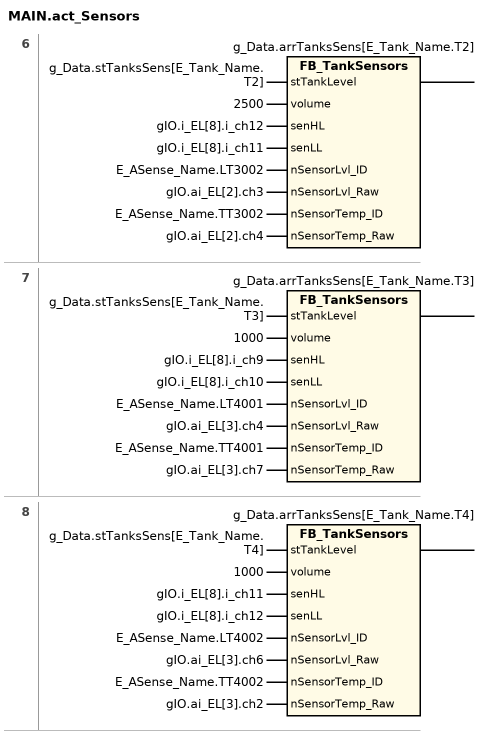
// NETWORK 6
g_Data.arrTanksSens[E_Tank_Name.T2](
    stTankLevel := g_Data.stTanksSens[E_Tank_Name.T2],
    volume := 2500,
    senHL := gIO.i_EL[8].i_ch12,
    senLL := gIO.i_EL[8].i_ch11,
    nSensorLvl_ID := E_ASense_Name.LT3002,
    nSensorLvl_Raw := gIO.ai_EL[2].ch3,
    nSensorTemp_ID := E_ASense_Name.TT3002,
    nSensorTemp_Raw := gIO.ai_EL[2].ch4); // FB_TankSensors

// NETWORK 7
g_Data.arrTanksSens[E_Tank_Name.T3](
    stTankLevel := g_Data.stTanksSens[E_Tank_Name.T3],
    volume := 1000,
    senHL := gIO.i_EL[8].i_ch9,
    senLL := gIO.i_EL[8].i_ch10,
    nSensorLvl_ID := E_ASense_Name.LT4001,
    nSensorLvl_Raw := gIO.ai_EL[3].ch4,
    nSensorTemp_ID := E_ASense_Name.TT4001,
    nSensorTemp_Raw := gIO.ai_EL[3].ch7); // FB_TankSensors

// NETWORK 8
g_Data.arrTanksSens[E_Tank_Name.T4](
    stTankLevel := g_Data.stTanksSens[E_Tank_Name.T4],
    volume := 1000,
    senHL := gIO.i_EL[8].i_ch11,
    senLL := gIO.i_EL[8].i_ch12,
    nSensorLvl_ID := E_ASense_Name.LT4002,
    nSensorLvl_Raw := gIO.ai_EL[3].ch6,
    nSensorTemp_ID := E_ASense_Name.TT4002,
    nSensorTemp_Raw := gIO.ai_EL[3].ch2); // FB_TankSensors
END_ACTION

ACTION act_SetAnalogSens_Test:
//set analog sensors setting only for the test. 
//Later this action should be deleted 
IF NOT bTesting THEN
	//Level
	g_AnalogSensor.stAnalogSensor[E_ASense_Name.LT1004].rawVal_Max:=14350;
	g_AnalogSensor.stAnalogSensor[E_ASense_Name.LT1004].rawVal_Min:=1270;
	g_AnalogSensor.stAnalogSensor[E_ASense_Name.LT1004].outVal_Max:=785;
	g_AnalogSensor.stAnalogSensor[E_ASense_Name.LT1004].outVal_Min:=0;
	g_AnalogSensor.stAnalogSensor[E_ASense_Name.LT1004].outOffset:=73;
	
	g_AnalogSensor.stAnalogSensor[E_ASense_Name.LT1003].rawVal_Max:=14350;
	g_AnalogSensor.stAnalogSensor[E_ASense_Name.LT1003].rawVal_Min:=1270;
	g_AnalogSensor.stAnalogSensor[E_ASense_Name.LT1003].outVal_Max:=785;
	g_AnalogSensor.stAnalogSensor[E_ASense_Name.LT1003].outVal_Min:=0;
	g_AnalogSensor.stAnalogSensor[E_ASense_Name.LT1003].outOffset:=73;
	
	g_AnalogSensor.stAnalogSensor[E_ASense_Name.LT1002].rawVal_Max:=14350;
	g_AnalogSensor.stAnalogSensor[E_ASense_Name.LT1002].rawVal_Min:=1270;
	g_AnalogSensor.stAnalogSensor[E_ASense_Name.LT1002].outVal_Max:=785;
	g_AnalogSensor.stAnalogSensor[E_ASense_Name.LT1002].outVal_Min:=0;
	g_AnalogSensor.stAnalogSensor[E_ASense_Name.LT1002].outOffset:=73;
	
	g_AnalogSensor.stAnalogSensor[E_ASense_Name.LT1001].rawVal_Max:=14350;
	g_AnalogSensor.stAnalogSensor[E_ASense_Name.LT1001].rawVal_Min:=1270;
	g_AnalogSensor.stAnalogSensor[E_ASense_Name.LT1001].outVal_Max:=785;
	g_AnalogSensor.stAnalogSensor[E_ASense_Name.LT1001].outVal_Min:=0;
	g_AnalogSensor.stAnalogSensor[E_ASense_Name.LT1001].outOffset:=73;
	
	//Flow
	g_AnalogSensor.stAnalogSensor[E_ASense_Name.FT1001].rawVal_Max:=10000;
	g_AnalogSensor.stAnalogSensor[E_ASense_Name.FT1001].rawVal_Min:=0;
	g_AnalogSensor.stAnalogSensor[E_ASense_Name.FT1001].outVal_Max:=306;
	g_AnalogSensor.stAnalogSensor[E_ASense_Name.FT1001].outVal_Min:=0;
	g_AnalogSensor.stAnalogSensor[E_ASense_Name.FT1001].outOffset:=0;
	
	g_AnalogSensor.stAnalogSensor[E_ASense_Name.FT1002].rawVal_Max:=10000;
	g_AnalogSensor.stAnalogSensor[E_ASense_Name.FT1002].rawVal_Min:=0;
	g_AnalogSensor.stAnalogSensor[E_ASense_Name.FT1002].outVal_Max:=306;
	g_AnalogSensor.stAnalogSensor[E_ASense_Name.FT1002].outVal_Min:=0;
	g_AnalogSensor.stAnalogSensor[E_ASense_Name.FT1002].outOffset:=0;
	
	////conductivity sensors
	g_AnalogSensor.stAnalogSensor[E_ASense_Name.CT1101].rawVal_Max:=14150;
	g_AnalogSensor.stAnalogSensor[E_ASense_Name.CT1101].rawVal_Min:=305;
	g_AnalogSensor.stAnalogSensor[E_ASense_Name.CT1101].outVal_Max:=14560;
	g_AnalogSensor.stAnalogSensor[E_ASense_Name.CT1101].outVal_Min:=346;
	g_AnalogSensor.stAnalogSensor[E_ASense_Name.CT1101].outOffset:=0;
	(*
	g_AnalogSensor.stAnalogSensor[E_ASense_Name.CT3101].rawVal_Max:=14150;
	g_AnalogSensor.stAnalogSensor[E_ASense_Name.CT3101].rawVal_Min:=305;
	g_AnalogSensor.stAnalogSensor[E_ASense_Name.CT3101].outVal_Max:=14560;
	g_AnalogSensor.stAnalogSensor[E_ASense_Name.CT3101].outVal_Min:=346;
	g_AnalogSensor.stAnalogSensor[E_ASense_Name.CT3101].outOffset:=0;
	*)
	//Temperature sensor
	g_AnalogSensor.stAnalogSensor[E_ASense_Name.TT1001].rawVal_Max:=7470;
	g_AnalogSensor.stAnalogSensor[E_ASense_Name.TT1001].rawVal_Min:=6400;
	g_AnalogSensor.stAnalogSensor[E_ASense_Name.TT1001].outVal_Max:=26;
	g_AnalogSensor.stAnalogSensor[E_ASense_Name.TT1001].outVal_Min:=20.9;
	g_AnalogSensor.stAnalogSensor[E_ASense_Name.TT1001].outOffset:=0;
	
	g_AnalogSensor.stAnalogSensor[E_ASense_Name.TT1002].rawVal_Max:=7470;
	g_AnalogSensor.stAnalogSensor[E_ASense_Name.TT1002].rawVal_Min:=6400;
	g_AnalogSensor.stAnalogSensor[E_ASense_Name.TT1002].outVal_Max:=26;
	g_AnalogSensor.stAnalogSensor[E_ASense_Name.TT1002].outVal_Min:=20.9;
	g_AnalogSensor.stAnalogSensor[E_ASense_Name.TT1002].outOffset:=0;
	
	g_AnalogSensor.stAnalogSensor[E_ASense_Name.TT1003].rawVal_Max:=7470;
	g_AnalogSensor.stAnalogSensor[E_ASense_Name.TT1003].rawVal_Min:=6400;
	g_AnalogSensor.stAnalogSensor[E_ASense_Name.TT1003].outVal_Max:=26;
	g_AnalogSensor.stAnalogSensor[E_ASense_Name.TT1003].outVal_Min:=20.9;
	g_AnalogSensor.stAnalogSensor[E_ASense_Name.TT1003].outOffset:=0;
	
	g_AnalogSensor.stAnalogSensor[E_ASense_Name.TT1004].rawVal_Max:=7470;
	g_AnalogSensor.stAnalogSensor[E_ASense_Name.TT1004].rawVal_Min:=6400;
	g_AnalogSensor.stAnalogSensor[E_ASense_Name.TT1004].outVal_Max:=26;
	g_AnalogSensor.stAnalogSensor[E_ASense_Name.TT1004].outVal_Min:=20.9;
	g_AnalogSensor.stAnalogSensor[E_ASense_Name.TT1004].outOffset:=0;
	
	g_AnalogSensor.stAnalogSensor[E_ASense_Name.TT1101].rawVal_Max:=7470;
	g_AnalogSensor.stAnalogSensor[E_ASense_Name.TT1101].rawVal_Min:=6400;
	g_AnalogSensor.stAnalogSensor[E_ASense_Name.TT1101].outVal_Max:=26;
	g_AnalogSensor.stAnalogSensor[E_ASense_Name.TT1101].outVal_Min:=20.9;
	g_AnalogSensor.stAnalogSensor[E_ASense_Name.TT1101].outOffset:=0;

	bTesting:=TRUE;
END_IF
END_ACTION

ACTION act_SetValves:
//Production tank
	//Tank1
	g_Data.arr_TankValves[1].valOutlet:=	E_Pis_Name.V3016;
	g_Data.arr_TankValves[1].valLine:=		E_Pis_Name.V3017;
	g_Data.arr_TankValves[1].valTriBlender:=E_Pis_Name.V3023;
	g_Data.arr_TankValves[1].valDrain:=		E_Pis_Name.V3024;
	g_Data.arr_TankValves[1].valCIP:=		E_Pis_Name.V3025;
	
	g_Data.arr_LineSourceValves[1].valTankA:=			E_Pis_Name.V3017;
	g_Data.arr_LineSourceValves[1].valTankB:=			E_Pis_Name.V3027;
	g_Data.arr_LineSourceValves[1].valTapWater:=		E_Pis_Name.V_Dummy_LSM_01;
	g_Data.arr_LineSourceValves[1].valTapWater_Drain:=	E_Pis_Name.V_Dummy_LSM_02;
	g_Data.arr_LineSourceValves[1].valTapWater_esle:=	E_Pis_Name.V_Dummy_LSM_05;
	g_Data.arr_LineSourceValves[1].valDrain:=			E_Pis_Name.V3018;
	g_Data.arr_LineSourceValves[1].valCIP:=				E_Pis_Name.V3019;
	g_Data.arr_LineSourceValves[1].valCIP_Sel:=			E_Pis_Name.V_Dummy_LSM_06;
	g_Data.arr_LineSourceValves[1].valBlockWater:=		E_Pis_Name.V_Dummy_LSM_03;
	g_Data.arr_LineSourceValves[1].valWaterSource:=		E_Pis_Name.V_Dummy_LSM_04;
	g_Data.arr_LineSourceValves[1].valWaterSource_Drain:=		E_Pis_Name.V_Dummy_LSM_07;
	
	g_Data.arr_TriBlenderSourceValves[1].valTankA:=				E_Pis_Name.V3023;
	g_Data.arr_TriBlenderSourceValves[1].valTankB:=				E_Pis_Name.V3028;
	g_Data.arr_TriBlenderSourceValves[1].valTapWater:=			E_Pis_Name.V_Dummy_TSM_01;
	g_Data.arr_TriBlenderSourceValves[1].valTapWater_Drain:=	E_Pis_Name.V_Dummy_TSM_02;
	g_Data.arr_TriBlenderSourceValves[1].valTapWater_esle:=		E_Pis_Name.V_Dummy_TSM_03;
	g_Data.arr_TriBlenderSourceValves[1].valDrain:=				E_Pis_Name.V3021;
	g_Data.arr_TriBlenderSourceValves[1].valCIP:=				E_Pis_Name.V3022;
	g_Data.arr_TriBlenderSourceValves[1].valCIP_Sel:=			E_Pis_Name.V3020;
	g_Data.arr_TriBlenderSourceValves[1].valBlockWater:=		E_Pis_Name.V3014;
	g_Data.arr_TriBlenderSourceValves[1].valWaterSource:=		E_Pis_Name.V3113;
	g_Data.arr_TriBlenderSourceValves[1].valWaterSource_Drain:=	E_Pis_Name.V2211;
	
	g_Data.arr_LineTargetValves[1].valTankA:=			E_Pis_Name.V_Dummy_01;//0;
	g_Data.arr_LineTargetValves[1].valTankB:=			E_Pis_Name.V_Dummy_02;//0;
	g_Data.arr_LineTargetValves[1].valDrain:=			E_Pis_Name.V_Dummy_03;//0;
	g_Data.arr_LineTargetValves[1].valCIP:=				E_Pis_Name.V_Dummy_04;//0;
	g_Data.arr_LineTargetValves[1].valTankA_Pipe:=		E_Pis_Name.V_Dummy_05;//0;
	g_Data.arr_LineTargetValves[1].valTankB_Pipe:=		E_Pis_Name.V_Dummy_06;//0;
	
	g_Data.arr_fbTriBlenderTargetValves[1].valTankA:=	E_Pis_Name.V3004;
	g_Data.arr_fbTriBlenderTargetValves[1].valTankB:=	E_Pis_Name.V3010;
	g_Data.arr_fbTriBlenderTargetValves[1].valDrain:=	E_Pis_Name.V3008;
	g_Data.arr_fbTriBlenderTargetValves[1].valCIP:=		E_Pis_Name.V3009;
	g_Data.arr_fbTriBlenderTargetValves[1].valTankA_Pipe:=		E_Pis_Name.v3041;
	g_Data.arr_fbTriBlenderTargetValves[1].valTankB_Pipe:=		E_Pis_Name.v3040;
	
	//Tank2
	g_Data.arr_TankValves[2].valOutlet:=	E_Pis_Name.V3015;
	g_Data.arr_TankValves[2].valLine:=		E_Pis_Name.V3027;
	g_Data.arr_TankValves[2].valTriBlender:=E_Pis_Name.V3028;
	g_Data.arr_TankValves[2].valDrain:=		E_Pis_Name.V3029;
	g_Data.arr_TankValves[2].valCIP:=		E_Pis_Name.V3030;
	
	g_Data.arr_LineSourceValves[2].valTankA:=			E_Pis_Name.V3017;
	g_Data.arr_LineSourceValves[2].valTankB:=			E_Pis_Name.V3027;
	g_Data.arr_LineSourceValves[2].valTapWater:=		E_Pis_Name.V_Dummy_LSM_01;
	g_Data.arr_LineSourceValves[2].valTapWater_Drain:=	E_Pis_Name.V_Dummy_LSM_02;
	g_Data.arr_LineSourceValves[2].valTapWater_esle:=	E_Pis_Name.V_Dummy_LSM_05;
	g_Data.arr_LineSourceValves[2].valDrain:=			E_Pis_Name.V3018;
	g_Data.arr_LineSourceValves[2].valCIP:=				E_Pis_Name.V3019;
	g_Data.arr_LineSourceValves[2].valCIP_Sel:=			E_Pis_Name.V_Dummy_LSM_06;
	g_Data.arr_LineSourceValves[2].valBlockWater:=		E_Pis_Name.V_Dummy_LSM_03;
	g_Data.arr_LineSourceValves[2].valWaterSource:=		E_Pis_Name.V_Dummy_LSM_04;
	g_Data.arr_LineSourceValves[2].valWaterSource_Drain:=		E_Pis_Name.V_Dummy_LSM_07;
	
	
	g_Data.arr_TriBlenderSourceValves[2].valTankA:=				E_Pis_Name.V3023;
	g_Data.arr_TriBlenderSourceValves[2].valTankB:=				E_Pis_Name.V3028;
	g_Data.arr_TriBlenderSourceValves[2].valTapWater:=			E_Pis_Name.V_Dummy_TSM_01;
	g_Data.arr_TriBlenderSourceValves[2].valTapWater_Drain:=	E_Pis_Name.V_Dummy_TSM_02;
	g_Data.arr_TriBlenderSourceValves[2].valTapWater_esle:=		E_Pis_Name.V_Dummy_TSM_03;
	g_Data.arr_TriBlenderSourceValves[2].valDrain:=				E_Pis_Name.V3021;
	g_Data.arr_TriBlenderSourceValves[2].valCIP:=				E_Pis_Name.V3022;
	g_Data.arr_TriBlenderSourceValves[2].valCIP_Sel:=			E_Pis_Name.V3020;
	g_Data.arr_TriBlenderSourceValves[2].valBlockWater:=		E_Pis_Name.V3014;
	g_Data.arr_TriBlenderSourceValves[2].valWaterSource:=		E_Pis_Name.V3113;
	g_Data.arr_TriBlenderSourceValves[2].valWaterSource_Drain:=	E_Pis_Name.V2211;
	
	g_Data.arr_LineTargetValves[2].valTankA:=			E_Pis_Name.V_Dummy_01;//0;
	g_Data.arr_LineTargetValves[2].valTankB:=			E_Pis_Name.V_Dummy_02;//0;
	g_Data.arr_LineTargetValves[2].valDrain:=			E_Pis_Name.V_Dummy_03;//0;
	g_Data.arr_LineTargetValves[2].valCIP:=				E_Pis_Name.V_Dummy_04;//0;
	g_Data.arr_LineTargetValves[2].valTankA_Pipe:=		E_Pis_Name.V_Dummy_05;//0;
	g_Data.arr_LineTargetValves[2].valTankB_Pipe:=		E_Pis_Name.V_Dummy_06;//0;	
	
	(*
	g_Data.arr_LineTargetValves[2].valTankA:=			E_Pis_Name.V_Dummy_07;//0;
	g_Data.arr_LineTargetValves[2].valTankB:=			E_Pis_Name.V_Dummy_08;//0;
	g_Data.arr_LineTargetValves[2].valDrain:=			E_Pis_Name.V_Dummy_09;//0;
	g_Data.arr_LineTargetValves[2].valCIP:=				E_Pis_Name.V_Dummy_10;//0;
	g_Data.arr_LineTargetValves[2].valTankA_Pipe:=		E_Pis_Name.V_Dummy_11;//0;
	g_Data.arr_LineTargetValves[2].valTankB_Pipe:=		E_Pis_Name.V_Dummy_12;//0;
	*)
	
	g_Data.arr_fbTriBlenderTargetValves[2].valTankA:=			E_Pis_Name.V3004;
	g_Data.arr_fbTriBlenderTargetValves[2].valTankB:=			E_Pis_Name.V3010;
	g_Data.arr_fbTriBlenderTargetValves[2].valDrain:=			E_Pis_Name.V3008;
	g_Data.arr_fbTriBlenderTargetValves[2].valCIP:=				E_Pis_Name.V3009;
	g_Data.arr_fbTriBlenderTargetValves[2].valTankA_Pipe:=		E_Pis_Name.V3041;
	g_Data.arr_fbTriBlenderTargetValves[2].valTankB_Pipe:=		E_Pis_Name.V3040;
	
	//Tank3
	g_Data.arr_TankValves[3].valOutlet:=	E_Pis_Name.V4016;
	g_Data.arr_TankValves[3].valLine:=		E_Pis_Name.V4017;
	g_Data.arr_TankValves[3].valTriBlender:=E_Pis_Name.V4023;
	g_Data.arr_TankValves[3].valDrain:=		E_Pis_Name.V4024;
	g_Data.arr_TankValves[3].valCIP:=		E_Pis_Name.V4025;
	
	g_Data.arr_LineSourceValves[3].valTankA:=			E_Pis_Name.V4017;
	g_Data.arr_LineSourceValves[3].valTankB:=			E_Pis_Name.V4027;
	g_Data.arr_LineSourceValves[3].valTapWater:=		E_Pis_Name.V2115;
	g_Data.arr_LineSourceValves[3].valTapWater_Drain:=	E_Pis_Name.V2117;
	g_Data.arr_LineSourceValves[3].valTapWater_esle:=	E_Pis_Name.V2116;
	g_Data.arr_LineSourceValves[3].valDrain:=			E_Pis_Name.V4018;
	g_Data.arr_LineSourceValves[3].valCIP:=				E_Pis_Name.V4019;
	g_Data.arr_LineSourceValves[3].valCIP_Sel:=			E_Pis_Name.V_Dummy_LSC_01;
	g_Data.arr_LineSourceValves[3].valBlockWater:=		E_Pis_Name.V_Dummy_LSC_02;
	g_Data.arr_LineSourceValves[3].valWaterSource:=		E_Pis_Name.V_Dummy_LSC_03;
	g_Data.arr_LineSourceValves[3].valWaterSource_Drain:=		E_Pis_Name.V_Dummy_LSC_04;
	
	g_Data.arr_TriBlenderSourceValves[3].valTankA:=				E_Pis_Name.V4023;
	g_Data.arr_TriBlenderSourceValves[3].valTankB:=				E_Pis_Name.V4028;
	g_Data.arr_TriBlenderSourceValves[3].valTapWater:=			E_Pis_Name.V2116;
	g_Data.arr_TriBlenderSourceValves[3].valTapWater_Drain:=	E_Pis_Name.V2117;
	g_Data.arr_TriBlenderSourceValves[3].valTapWater_esle:=		E_Pis_Name.V2115;
	g_Data.arr_TriBlenderSourceValves[3].valDrain:=				E_Pis_Name.V4021;
	g_Data.arr_TriBlenderSourceValves[3].valCIP:=				E_Pis_Name.V4022;
	g_Data.arr_TriBlenderSourceValves[3].valCIP_Sel:=			E_Pis_Name.V4020;
	g_Data.arr_TriBlenderSourceValves[3].valBlockWater:=		E_Pis_Name.V4014;
	g_Data.arr_TriBlenderSourceValves[3].valWaterSource:=		E_Pis_Name.V2114;
	g_Data.arr_TriBlenderSourceValves[3].valWaterSource_Drain:=	E_Pis_Name.V2112;
	
	g_Data.arr_LineTargetValves[3].valTankA:=	E_Pis_Name.V4034;
	g_Data.arr_LineTargetValves[3].valTankB:=	E_Pis_Name.V4033;
	g_Data.arr_LineTargetValves[3].valDrain:=	E_Pis_Name.V4035;
	g_Data.arr_LineTargetValves[3].valCIP:=		E_Pis_Name.V4036;
	g_Data.arr_LineTargetValves[3].valTankA_Pipe:=		E_Pis_Name.V4041;
	g_Data.arr_LineTargetValves[3].valTankB_Pipe:=		E_Pis_Name.V4040;
	
	g_Data.arr_fbTriBlenderTargetValves[3].valTankA:=	E_Pis_Name.V4004;
	g_Data.arr_fbTriBlenderTargetValves[3].valTankB:=	E_Pis_Name.V4010;
	g_Data.arr_fbTriBlenderTargetValves[3].valDrain:=	E_Pis_Name.V4008;
	g_Data.arr_fbTriBlenderTargetValves[3].valCIP:=		E_Pis_Name.V4009;
	g_Data.arr_fbTriBlenderTargetValves[3].valTankA_Pipe:=		E_Pis_Name.V4041;
	g_Data.arr_fbTriBlenderTargetValves[3].valTankB_Pipe:=		E_Pis_Name.V4040;
	
	//Tank4
	g_Data.arr_TankValves[4].valOutlet:=	E_Pis_Name.V4015;
	g_Data.arr_TankValves[4].valLine:=		E_Pis_Name.V4027;
	g_Data.arr_TankValves[4].valTriBlender:=E_Pis_Name.V4028;
	g_Data.arr_TankValves[4].valDrain:=		E_Pis_Name.V4029;
	g_Data.arr_TankValves[4].valCIP:=		E_Pis_Name.V4030;
	
	g_Data.arr_LineSourceValves[4].valTankA:=			E_Pis_Name.V4017;
	g_Data.arr_LineSourceValves[4].valTankB:=			E_Pis_Name.V4027;
	g_Data.arr_LineSourceValves[4].valTapWater:=		E_Pis_Name.V2115;
	g_Data.arr_LineSourceValves[4].valTapWater_Drain:=	E_Pis_Name.V2117;
	g_Data.arr_LineSourceValves[4].valTapWater_esle:=	E_Pis_Name.V2116;
	g_Data.arr_LineSourceValves[4].valDrain:=			E_Pis_Name.V4018;
	g_Data.arr_LineSourceValves[4].valCIP:=				E_Pis_Name.V4019;
	g_Data.arr_LineSourceValves[4].valCIP_Sel:=			E_Pis_Name.V_Dummy_LSC_01;
	g_Data.arr_LineSourceValves[4].valBlockWater:=		E_Pis_Name.V_Dummy_LSC_02;
	g_Data.arr_LineSourceValves[4].valWaterSource:=		E_Pis_Name.V_Dummy_LSC_03;
	g_Data.arr_LineSourceValves[4].valWaterSource_Drain:=		E_Pis_Name.V_Dummy_LSC_04;
	
	g_Data.arr_TriBlenderSourceValves[4].valTankA:=				E_Pis_Name.V4023;
	g_Data.arr_TriBlenderSourceValves[4].valTankB:=				E_Pis_Name.V4028;
	g_Data.arr_TriBlenderSourceValves[4].valTapWater:=			E_Pis_Name.V2116;
	g_Data.arr_TriBlenderSourceValves[4].valTapWater_Drain:=	E_Pis_Name.V2117;
	g_Data.arr_TriBlenderSourceValves[4].valTapWater_esle:=		E_Pis_Name.V2115;
	g_Data.arr_TriBlenderSourceValves[4].valDrain:=				E_Pis_Name.V4021;
	g_Data.arr_TriBlenderSourceValves[4].valCIP:=				E_Pis_Name.V4022;
	g_Data.arr_TriBlenderSourceValves[4].valCIP_Sel:=			E_Pis_Name.V4020;
	g_Data.arr_TriBlenderSourceValves[4].valBlockWater:=		E_Pis_Name.V4014;
	g_Data.arr_TriBlenderSourceValves[4].valWaterSource:=		E_Pis_Name.V2114;
	g_Data.arr_TriBlenderSourceValves[4].valWaterSource_Drain:=	E_Pis_Name.V2112;
	
	g_Data.arr_LineTargetValves[4].valTankA:=	E_Pis_Name.V4034;
	g_Data.arr_LineTargetValves[4].valTankB:=	E_Pis_Name.V4033;
	g_Data.arr_LineTargetValves[4].valDrain:=	E_Pis_Name.V4035;
	g_Data.arr_LineTargetValves[4].valCIP:=		E_Pis_Name.V4036;
	g_Data.arr_LineTargetValves[4].valTankA_Pipe:=		E_Pis_Name.V4041;
	g_Data.arr_LineTargetValves[4].valTankB_Pipe:=		E_Pis_Name.V4040;
	
	g_Data.arr_fbTriBlenderTargetValves[4].valTankA:=	E_Pis_Name.V4004;
	g_Data.arr_fbTriBlenderTargetValves[4].valTankB:=	E_Pis_Name.V4010;
	g_Data.arr_fbTriBlenderTargetValves[4].valDrain:=	E_Pis_Name.V4008;
	g_Data.arr_fbTriBlenderTargetValves[4].valCIP:=		E_Pis_Name.V4009;
	g_Data.arr_fbTriBlenderTargetValves[4].valTankA_Pipe:=		E_Pis_Name.V4041;
	g_Data.arr_fbTriBlenderTargetValves[4].valTankB_Pipe:=		E_Pis_Name.V4040;
END_ACTION

METHOD m_TankConus_Level_Calculation : REAL
VAR_INPUT
	raw: REAL;

END_VAR
VAR
	kConus: REAL:=0.00000002149 ;
END_VAR
IF raw<1230 THEN;
	//m_TankConus_Level_Calculation:=kConus*raw^3;
ELSE;
	m_TankConus_Level_Calculation:=raw;
END_IF
END_METHOD

METHOD mElementList_SetName : BOOL
VAR_INPUT
END_VAR

VAR
	eASense_Name: E_ASense_Name;
	eProcCntrl: E_ProcessControl_Name;
END_VAR
FOR eASense_Name:=0 TO E_ASense_Name.last DO
	arAnalogSensorNameList[eASense_Name]:=TO_STRING(eASense_Name);
END_FOR

FOR eProcCntrl:=0 TO E_ProcessControl_Name.eProcCntrl_Last DO
	arr_ProcCntrl_NameList[eProcCntrl]:=TO_STRING(eProcCntrl);
	g_ProcControl.arr_stProcCntrl[eProcCntrl].idName:=TO_STRING(eProcCntrl);
END_FOR
END_METHOD

END_PROGRAM

// ---- 03 Project/40 Misc/FB_OpenClose_Vlave.TcPOU
FUNCTION_BLOCK FB_OpenClose_Vlave
VAR_INPUT
	val_AfterPump	: E_Pis_Name;
	Pump_ID			: E_Pump_List:=E_Pump_List.eNotSelected;
END_VAR
VAR_OUTPUT
END_VAR
VAR
	stPist	: REFERENCE TO ST_Piston;
	stPump	: REFERENCE TO ST_Pump	;
	bOneTime	:	BOOL	;
END_VAR

act_SetReference();

IF (stPump.bRun_Auto OR stPump.bRun_Man) THEN
	bOneTime:=FALSE;
	IF NOT stPist.st_Open THEN
		stPist.req_Open:=TRUE;
	END_IF
ELSE
	IF NOT stPist.st_Close AND NOT bOneTime THEN
		stPist.req_Close:=TRUE;
		bOneTime:=TRUE;
	END_IF
END_IF

ACTION act_SetReference:
stPist REF= stPis[val_AfterPump];
stPump REF= g_Pump.arr_st_Pump[Pump_ID];
END_ACTION

END_FUNCTION_BLOCK

// ---- 00 Library/00-General/TimeAndDate/prg_RealClock.TcPOU
PROGRAM prg_RealClock
VAR

(* Real Time Clock *)
(*	dtRealTime				: DATE_AND_TIME;
	sRealTime				: STRING[22];	
	stSystemTime			: TimeStruct;
	stSystemTime_Empty		: TimeStruct;
	sTime					: STRING[20];
	sDate					: STRING[20];
	sTimeWithMicroSec		: STRING[40];*)

	syncTimer 	: TON;
	fbGetLocalTime 	: NT_GetTime;
	fbRTC_EX2 	: RTC_EX2;
	presetTime 	: TimeStruct;
	syncTrigger 	: F_TRIG;
	bBusy 		: BOOL;
	bError 		: BOOL;
	nErrID 		: UDINT;
	temp1: DATE;
	temp2: TOD;
	NetId :STRING :='';
	bValid_RTCEX2 	: BOOL;
	nMicroseconds 	: DWORD;
	r_trigTrigger: R_TRIG;
	sRealTime_Date	 :STRING(25);
	
	bStartTime: BOOL;
	stStart: TimeStruct;
	sDelta: STRING;
	ton_OneMinuteCount: TON;
END_VAR

(*--------->Set Plc Clock<----------------*)

dtRealTime:=SYSTEMTIME_TO_DT(stSystemTime);
sRealTime:= DT_TO_STRING(dtRealTime);
sRealTime_Date:= DT_TO_STRING(dtRealTime);
sRealTime_Date:=right(sRealTime_Date,19);
temp1:=DT_TO_DATE(dtRealTime);
temp2:=DT_TO_TOD(dtRealTime);
sDate:=DATE_TO_STRING(temp1);
sDate:=DELETE(sDate,2,1);


sTime:=TOD_TO_STRING(temp2);
sTime:=DELETE(sTime,4,1);

sDateTime:=CONCAT(sDate,' ');
sDateTime:=CONCAT(sDateTime,sTime);

sTimeWithMicroSec:=CONCAT(sTime,'.');
sTimeWithMicroSec:=CONCAT(sTimeWithMicroSec,DWORD_TO_STRING(nMicroseconds));




	syncTimer(IN:=NOT SyncTimer.Q , PT:=T#100ms , Q=> , ET=> );
(*r_trigTrigger(CLK:=q_Trigger);*)
	fbGetLocalTime(
		NETID:='' ,
		START:=syncTimer.Q,
		(*START:=r_trigTrigger.Q,*)
		TMOUT:=T#5s ,
		BUSY=>bBusy ,
		ERR=>bError ,
		ERRID=>nErrId ,
		TIMESTR=>presetTime );

	(*syncTrigger(CLK:=NOT bBusy*)
	syncTrigger(CLK:= bBusy
					 AND NOT bError , Q=> );
	fbRTC_EX2(
		EN:=syncTrigger.Q ,
		PDT:=presetTime ,
		PMICRO:=0 ,
		Q=>bValid_RTCEX2 ,
		CDT=>stSystemTime ,
		CMICRO=>nMicroseconds );
		
act_TestDelta();	

ton_OneMinuteCount(PT:=T#1m, IN:=NOT ton_OneMinuteCount.Q);

ACTION act_TestDelta:
IF bStartTime THEN;
	bStartTime:=FALSE;
	stStart:=stSystemTime;
END_IF

sDelta:= m_DeltaTime(stStartTime:=stStart);
END_ACTION

METHOD m_DeltaTime : STRING
VAR_INPUT
	stStartTime  : TimeStruct;
END_VAR
VAR
	tDelta: TIME;
	dtDelta: DATE_AND_TIME;
	todDelta: TOD;


END_VAR
tDelta:=TO_TIME(SYSTEMTIME_TO_DT(stSystemTime)-SYSTEMTIME_TO_DT(stStartTime));

m_DeltaTime:=mTime_to_String_HMI(tInputTime:=tDelta,iSecondDisplay:=FALSE);

(*old
todDelta:=TIME_TO_TOD(tDelta);
m_DeltaTime:=TOD_TO_STRING(todDelta);
m_DeltaTime:=DELETE(m_DeltaTime,4,1);
//dtDelta:=TO_DT(SYSTEMTIME_TO_DT(stSystemTime)-SYSTEMTIME_TO_DT(stStartTime));
//m_DeltaTime:=TIME_TO_STRING(dtDelta);
*)
END_METHOD

METHOD mTime_to_String_HMI : STRING
VAR_INPUT
    tInputTime 		: TIME; // TIME type, stored internally as LTIME (ms)
	iSecondDisplay	: BOOL;
END_VAR
VAR
    nTotalSeconds : UDINT;
    nTotalHours : UDINT;
    nMinutes : UDINT;
    nSeconds : UDINT;
    sFormatted : STRING(20);
END_VAR
// Convert TIME to total seconds
nTotalSeconds := TO_UDINT(tInputTime) / 1000;

// Extract minutes and seconds
nMinutes := nTotalSeconds / 60;
nSeconds := nTotalSeconds MOD 60;

// Convert to total hours
nTotalHours := nMinutes / 60;
nMinutes := nMinutes MOD 60;

// Format output as HHHH:MM:SS (e.g., 0123:45:56)
sFormatted := CONCAT(UDINT_TO_STRING(nTotalHours),'h:');
IF nMinutes < 10 THEN
    sFormatted := CONCAT(sFormatted, '0');
END_IF
sFormatted := CONCAT(sFormatted, UDINT_TO_STRING(nMinutes));
sFormatted := CONCAT(sFormatted, 'm');

IF iSecondDisplay THEN;
	sFormatted := CONCAT(sFormatted, ':');
	IF nSeconds < 10 THEN
		sFormatted := CONCAT(sFormatted, '0');
	END_IF
	sFormatted := CONCAT(sFormatted, UDINT_TO_STRING(nSeconds));
	sFormatted := CONCAT(sFormatted, 's');	
END_IF

// Return formatted string
mTime_to_String_HMI := sFormatted;
END_METHOD

END_PROGRAM

// ---- 01 Instance/01 Piston/prg_Piston.TcPOU
PROGRAM prg_Piston
VAR
	fbPiston: FB_Piston;
	stPiston: ST_Piston;

	bPis_Next_P: BOOL;
	bPis_Next_N: BOOL;

	

	
	TON_0: TON;
	TON_1: TON;
	TON_2: TON;
	TON_3: TON;
	TON_4: TON;
	TON_5: TON;	
	i: INT;
END_VAR

act_InterLock();
act_Call_list_TanksMarinade();
act_Call_list_TanksColor();
act_Call_list_TanksCoolant();
act_Call_List_LineSource();
act_Call_List_LineTarget();
act_Call_list_CIP_SourceNTarget();
act_Call_list_CIP_Client();
act_Call_list_CIP_Tanks();
act_Call_list_Water();
act_Call_list_TriBlender_Selector();


IF bPis_Next_P THEN;
	m_Get_Next_P(iSel:=iPis_sel);
	bPis_Next_P:=FALSE;
END_IF

IF bPis_Next_N THEN;
	m_Get_Next_N(iSel:=iPis_sel);
	bPis_Next_N:=FALSE;
END_IF

FOR i:=0 TO E_Pis_Name.last DO
	ePisNameList:=i;
	arPisNameList[i]:=TO_STRING(ePisNameList);
END_FOR

ACTION act_Call_list_CIP_Client:
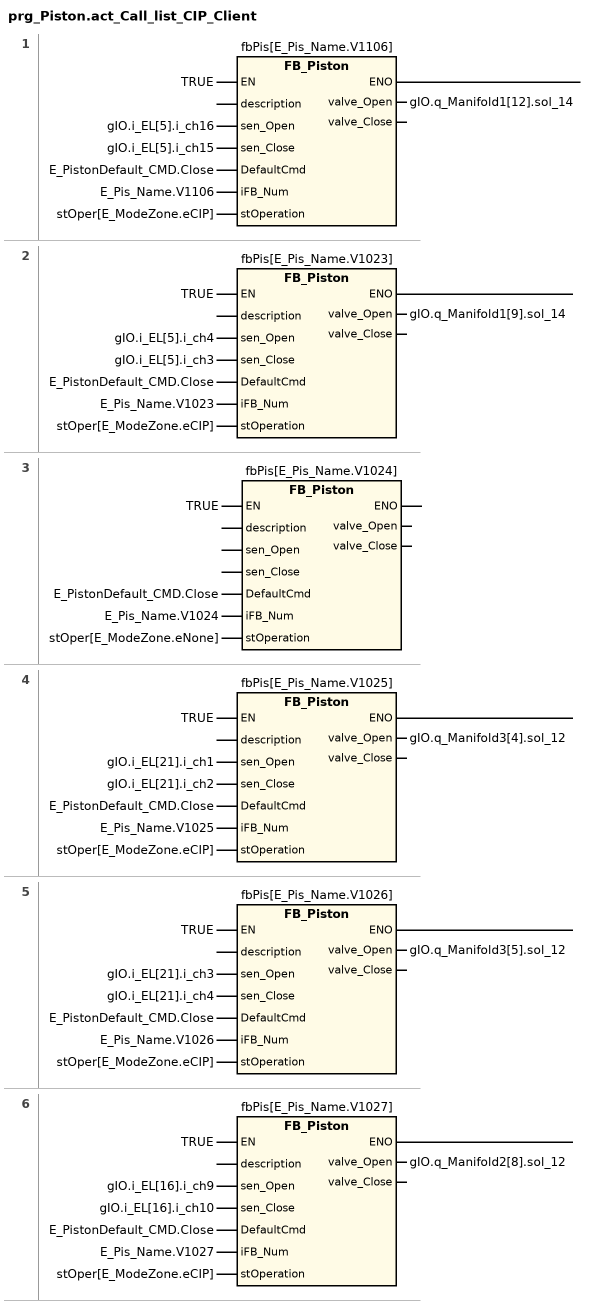
// NETWORK 1
fbPis[E_Pis_Name.V1106](
    sen_Open := gIO.i_EL[5].i_ch16,
    sen_Close := gIO.i_EL[5].i_ch15,
    DefaultCmd := E_PistonDefault_CMD.Close,
    iFB_Num := E_Pis_Name.V1106,
    stOperation := stOper[E_ModeZone.eCIP],
    valve_Open => gIO.q_Manifold1[12].sol_14); // FB_Piston

// NETWORK 2
fbPis[E_Pis_Name.V1023](
    sen_Open := gIO.i_EL[5].i_ch4,
    sen_Close := gIO.i_EL[5].i_ch3,
    DefaultCmd := E_PistonDefault_CMD.Close,
    iFB_Num := E_Pis_Name.V1023,
    stOperation := stOper[E_ModeZone.eCIP],
    valve_Open => gIO.q_Manifold1[9].sol_14); // FB_Piston

// NETWORK 3
fbPis[E_Pis_Name.V1024](
    DefaultCmd := E_PistonDefault_CMD.Close,
    iFB_Num := E_Pis_Name.V1024,
    stOperation := stOper[E_ModeZone.eNone]); // FB_Piston

// NETWORK 4
fbPis[E_Pis_Name.V1025](
    sen_Open := gIO.i_EL[21].i_ch1,
    sen_Close := gIO.i_EL[21].i_ch2,
    DefaultCmd := E_PistonDefault_CMD.Close,
    iFB_Num := E_Pis_Name.V1025,
    stOperation := stOper[E_ModeZone.eCIP],
    valve_Open => gIO.q_Manifold3[4].sol_12); // FB_Piston

// NETWORK 5
fbPis[E_Pis_Name.V1026](
    sen_Open := gIO.i_EL[21].i_ch3,
    sen_Close := gIO.i_EL[21].i_ch4,
    DefaultCmd := E_PistonDefault_CMD.Close,
    iFB_Num := E_Pis_Name.V1026,
    stOperation := stOper[E_ModeZone.eCIP],
    valve_Open => gIO.q_Manifold3[5].sol_12); // FB_Piston

// NETWORK 6
fbPis[E_Pis_Name.V1027](
    sen_Open := gIO.i_EL[16].i_ch9,
    sen_Close := gIO.i_EL[16].i_ch10,
    DefaultCmd := E_PistonDefault_CMD.Close,
    iFB_Num := E_Pis_Name.V1027,
    stOperation := stOper[E_ModeZone.eCIP],
    valve_Open => gIO.q_Manifold2[8].sol_12); // FB_Piston

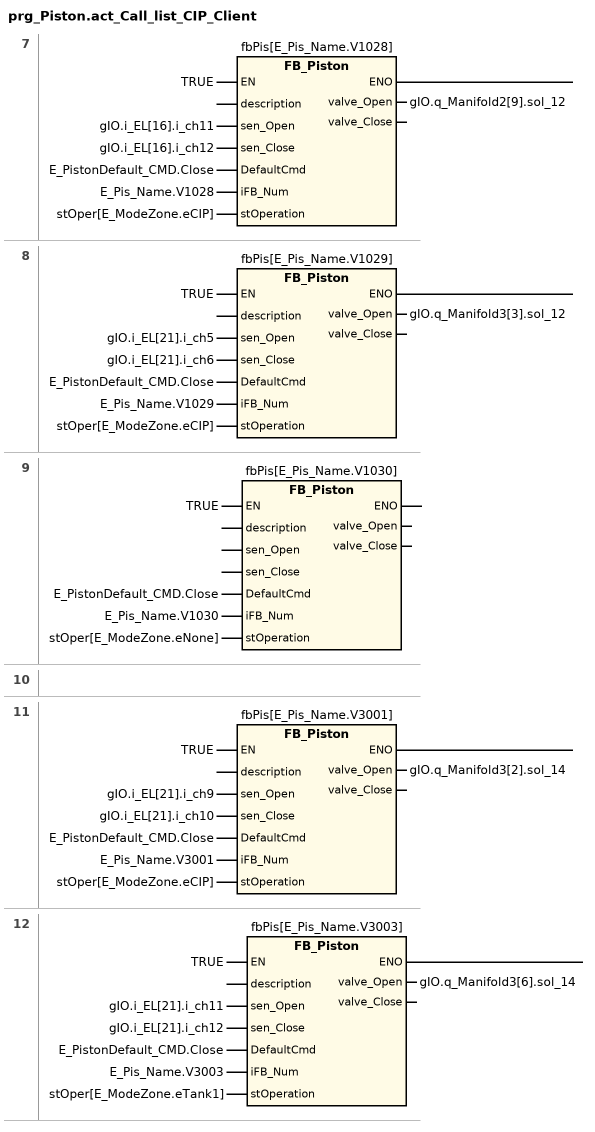
// NETWORK 7
fbPis[E_Pis_Name.V1028](
    sen_Open := gIO.i_EL[16].i_ch11,
    sen_Close := gIO.i_EL[16].i_ch12,
    DefaultCmd := E_PistonDefault_CMD.Close,
    iFB_Num := E_Pis_Name.V1028,
    stOperation := stOper[E_ModeZone.eCIP],
    valve_Open => gIO.q_Manifold2[9].sol_12); // FB_Piston

// NETWORK 8
fbPis[E_Pis_Name.V1029](
    sen_Open := gIO.i_EL[21].i_ch5,
    sen_Close := gIO.i_EL[21].i_ch6,
    DefaultCmd := E_PistonDefault_CMD.Close,
    iFB_Num := E_Pis_Name.V1029,
    stOperation := stOper[E_ModeZone.eCIP],
    valve_Open => gIO.q_Manifold3[3].sol_12); // FB_Piston

// NETWORK 9
fbPis[E_Pis_Name.V1030](
    DefaultCmd := E_PistonDefault_CMD.Close,
    iFB_Num := E_Pis_Name.V1030,
    stOperation := stOper[E_ModeZone.eNone]); // FB_Piston

// NETWORK 10

// NETWORK 11
fbPis[E_Pis_Name.V3001](
    sen_Open := gIO.i_EL[21].i_ch9,
    sen_Close := gIO.i_EL[21].i_ch10,
    DefaultCmd := E_PistonDefault_CMD.Close,
    iFB_Num := E_Pis_Name.V3001,
    stOperation := stOper[E_ModeZone.eCIP],
    valve_Open => gIO.q_Manifold3[2].sol_14); // FB_Piston

// NETWORK 12
fbPis[E_Pis_Name.V3003](
    sen_Open := gIO.i_EL[21].i_ch11,
    sen_Close := gIO.i_EL[21].i_ch12,
    DefaultCmd := E_PistonDefault_CMD.Close,
    iFB_Num := E_Pis_Name.V3003,
    stOperation := stOper[E_ModeZone.eTank1],
    valve_Open => gIO.q_Manifold3[6].sol_14); // FB_Piston

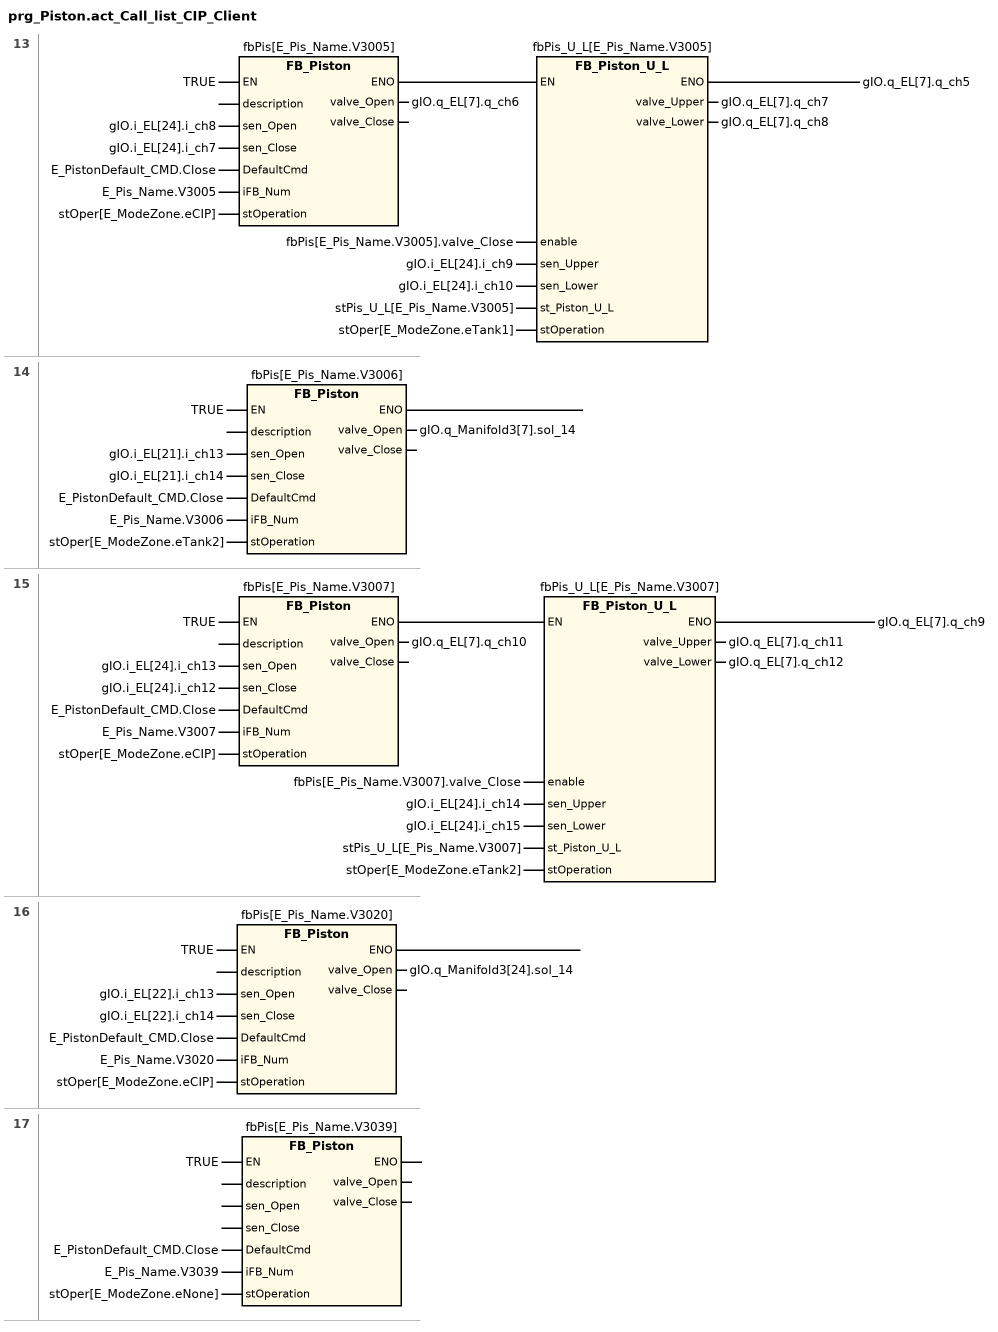
// NETWORK 13
fbPis[E_Pis_Name.V3005](
    sen_Open := gIO.i_EL[24].i_ch8,
    sen_Close := gIO.i_EL[24].i_ch7,
    DefaultCmd := E_PistonDefault_CMD.Close,
    iFB_Num := E_Pis_Name.V3005,
    stOperation := stOper[E_ModeZone.eCIP],
    valve_Open => gIO.q_EL[7].q_ch6); // FB_Piston
fbPis_U_L[E_Pis_Name.V3005](
    enable := fbPis[E_Pis_Name.V3005].valve_Close,
    sen_Upper := gIO.i_EL[24].i_ch9,
    sen_Lower := gIO.i_EL[24].i_ch10,
    st_Piston_U_L := stPis_U_L[E_Pis_Name.V3005],
    stOperation := stOper[E_ModeZone.eTank1],
    valve_Upper => gIO.q_EL[7].q_ch7,
    valve_Lower => gIO.q_EL[7].q_ch8); // FB_Piston_U_L
gIO.q_EL[7].q_ch5 := TRUE;

// NETWORK 14
fbPis[E_Pis_Name.V3006](
    sen_Open := gIO.i_EL[21].i_ch13,
    sen_Close := gIO.i_EL[21].i_ch14,
    DefaultCmd := E_PistonDefault_CMD.Close,
    iFB_Num := E_Pis_Name.V3006,
    stOperation := stOper[E_ModeZone.eTank2],
    valve_Open => gIO.q_Manifold3[7].sol_14); // FB_Piston

// NETWORK 15
fbPis[E_Pis_Name.V3007](
    sen_Open := gIO.i_EL[24].i_ch13,
    sen_Close := gIO.i_EL[24].i_ch12,
    DefaultCmd := E_PistonDefault_CMD.Close,
    iFB_Num := E_Pis_Name.V3007,
    stOperation := stOper[E_ModeZone.eCIP],
    valve_Open => gIO.q_EL[7].q_ch10); // FB_Piston
fbPis_U_L[E_Pis_Name.V3007](
    enable := fbPis[E_Pis_Name.V3007].valve_Close,
    sen_Upper := gIO.i_EL[24].i_ch14,
    sen_Lower := gIO.i_EL[24].i_ch15,
    st_Piston_U_L := stPis_U_L[E_Pis_Name.V3007],
    stOperation := stOper[E_ModeZone.eTank2],
    valve_Upper => gIO.q_EL[7].q_ch11,
    valve_Lower => gIO.q_EL[7].q_ch12); // FB_Piston_U_L
gIO.q_EL[7].q_ch9 := TRUE;

// NETWORK 16
fbPis[E_Pis_Name.V3020](
    sen_Open := gIO.i_EL[22].i_ch13,
    sen_Close := gIO.i_EL[22].i_ch14,
    DefaultCmd := E_PistonDefault_CMD.Close,
    iFB_Num := E_Pis_Name.V3020,
    stOperation := stOper[E_ModeZone.eCIP],
    valve_Open => gIO.q_Manifold3[24].sol_14); // FB_Piston

// NETWORK 17
fbPis[E_Pis_Name.V3039](
    DefaultCmd := E_PistonDefault_CMD.Close,
    iFB_Num := E_Pis_Name.V3039,
    stOperation := stOper[E_ModeZone.eNone]); // FB_Piston

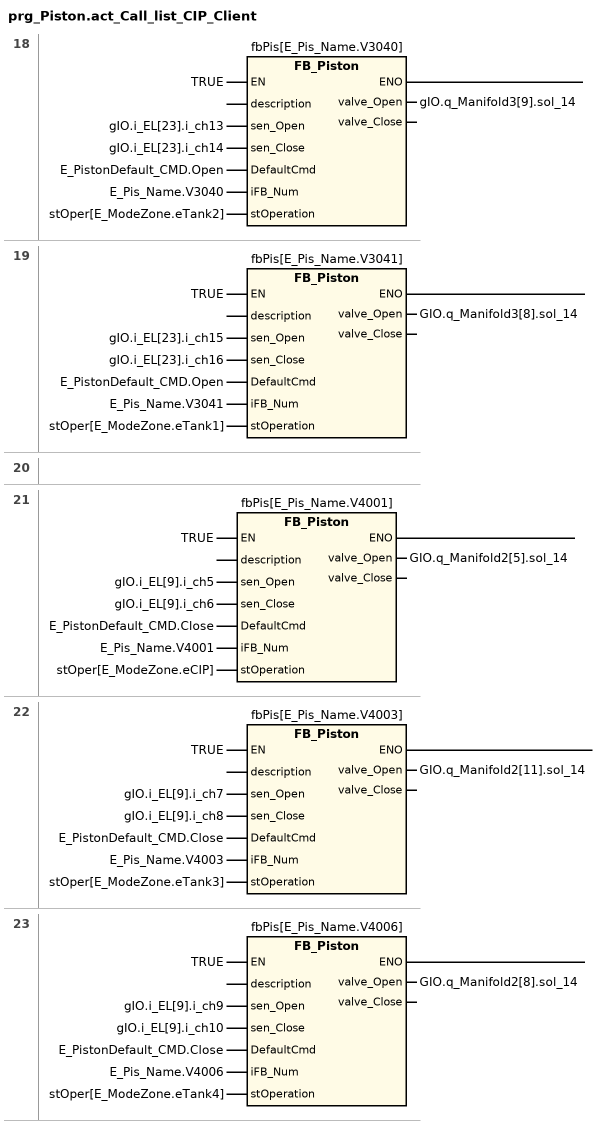
// NETWORK 18
fbPis[E_Pis_Name.V3040](
    sen_Open := gIO.i_EL[23].i_ch13,
    sen_Close := gIO.i_EL[23].i_ch14,
    DefaultCmd := E_PistonDefault_CMD.Open,
    iFB_Num := E_Pis_Name.V3040,
    stOperation := stOper[E_ModeZone.eTank2],
    valve_Open => gIO.q_Manifold3[9].sol_14); // FB_Piston

// NETWORK 19
fbPis[E_Pis_Name.V3041](
    sen_Open := gIO.i_EL[23].i_ch15,
    sen_Close := gIO.i_EL[23].i_ch16,
    DefaultCmd := E_PistonDefault_CMD.Open,
    iFB_Num := E_Pis_Name.V3041,
    stOperation := stOper[E_ModeZone.eTank1],
    valve_Open => GIO.q_Manifold3[8].sol_14); // FB_Piston

// NETWORK 20

// NETWORK 21
fbPis[E_Pis_Name.V4001](
    sen_Open := gIO.i_EL[9].i_ch5,
    sen_Close := gIO.i_EL[9].i_ch6,
    DefaultCmd := E_PistonDefault_CMD.Close,
    iFB_Num := E_Pis_Name.V4001,
    stOperation := stOper[E_ModeZone.eCIP],
    valve_Open => GIO.q_Manifold2[5].sol_14); // FB_Piston

// NETWORK 22
fbPis[E_Pis_Name.V4003](
    sen_Open := gIO.i_EL[9].i_ch7,
    sen_Close := gIO.i_EL[9].i_ch8,
    DefaultCmd := E_PistonDefault_CMD.Close,
    iFB_Num := E_Pis_Name.V4003,
    stOperation := stOper[E_ModeZone.eTank3],
    valve_Open => GIO.q_Manifold2[11].sol_14); // FB_Piston

// NETWORK 23
fbPis[E_Pis_Name.V4006](
    sen_Open := gIO.i_EL[9].i_ch9,
    sen_Close := gIO.i_EL[9].i_ch10,
    DefaultCmd := E_PistonDefault_CMD.Close,
    iFB_Num := E_Pis_Name.V4006,
    stOperation := stOper[E_ModeZone.eTank4],
    valve_Open => GIO.q_Manifold2[8].sol_14); // FB_Piston

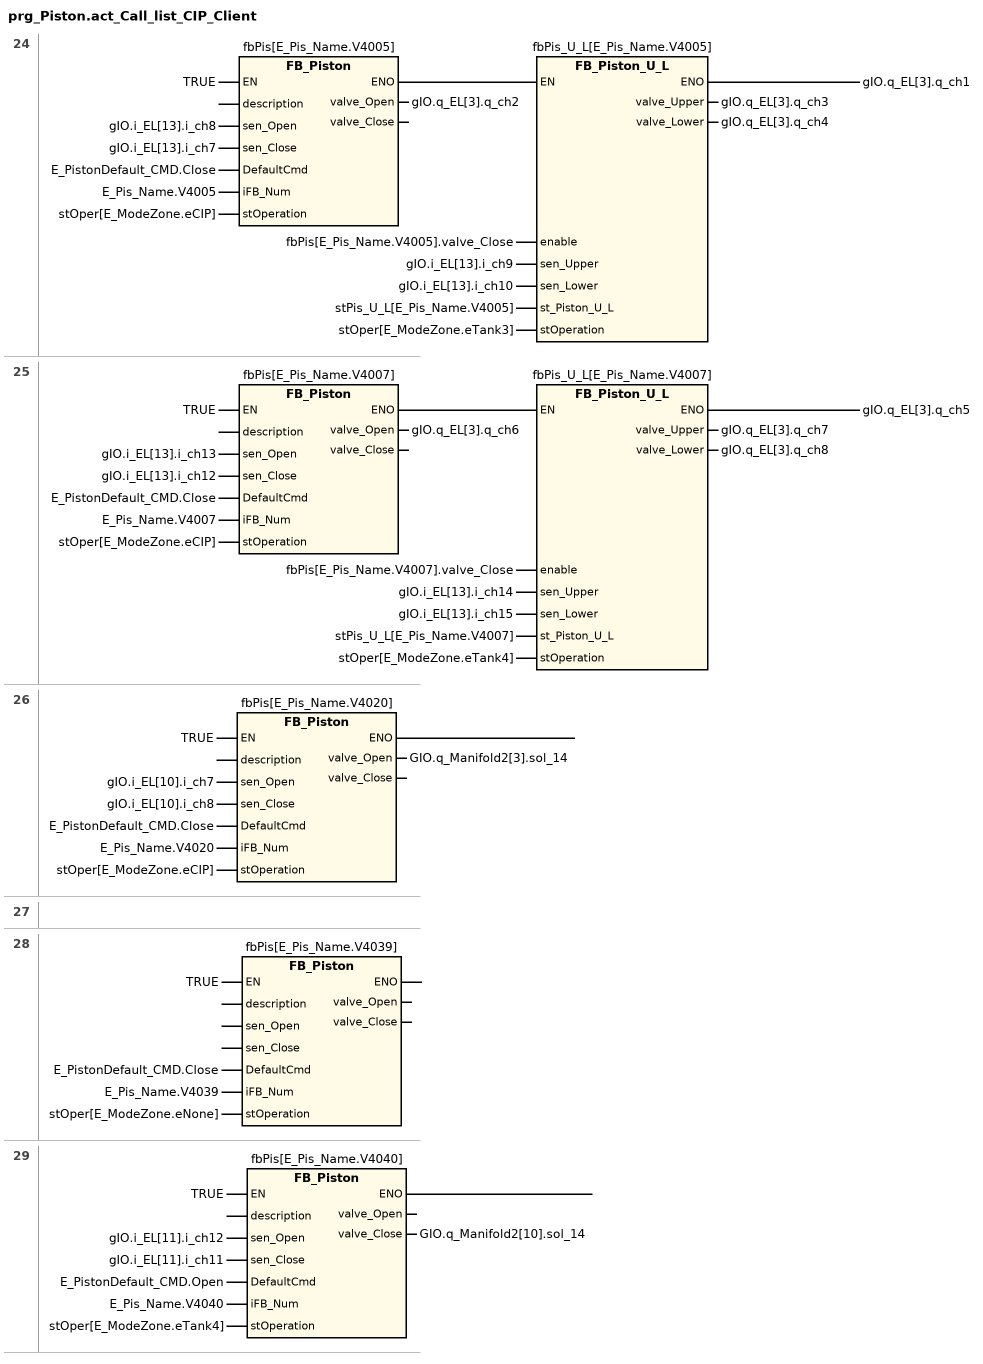
// NETWORK 24
fbPis[E_Pis_Name.V4005](
    sen_Open := gIO.i_EL[13].i_ch8,
    sen_Close := gIO.i_EL[13].i_ch7,
    DefaultCmd := E_PistonDefault_CMD.Close,
    iFB_Num := E_Pis_Name.V4005,
    stOperation := stOper[E_ModeZone.eCIP],
    valve_Open => gIO.q_EL[3].q_ch2); // FB_Piston
fbPis_U_L[E_Pis_Name.V4005](
    enable := fbPis[E_Pis_Name.V4005].valve_Close,
    sen_Upper := gIO.i_EL[13].i_ch9,
    sen_Lower := gIO.i_EL[13].i_ch10,
    st_Piston_U_L := stPis_U_L[E_Pis_Name.V4005],
    stOperation := stOper[E_ModeZone.eTank3],
    valve_Upper => gIO.q_EL[3].q_ch3,
    valve_Lower => gIO.q_EL[3].q_ch4); // FB_Piston_U_L
gIO.q_EL[3].q_ch1 := TRUE;

// NETWORK 25
fbPis[E_Pis_Name.V4007](
    sen_Open := gIO.i_EL[13].i_ch13,
    sen_Close := gIO.i_EL[13].i_ch12,
    DefaultCmd := E_PistonDefault_CMD.Close,
    iFB_Num := E_Pis_Name.V4007,
    stOperation := stOper[E_ModeZone.eCIP],
    valve_Open => gIO.q_EL[3].q_ch6); // FB_Piston
fbPis_U_L[E_Pis_Name.V4007](
    enable := fbPis[E_Pis_Name.V4007].valve_Close,
    sen_Upper := gIO.i_EL[13].i_ch14,
    sen_Lower := gIO.i_EL[13].i_ch15,
    st_Piston_U_L := stPis_U_L[E_Pis_Name.V4007],
    stOperation := stOper[E_ModeZone.eTank4],
    valve_Upper => gIO.q_EL[3].q_ch7,
    valve_Lower => gIO.q_EL[3].q_ch8); // FB_Piston_U_L
gIO.q_EL[3].q_ch5 := TRUE;

// NETWORK 26
fbPis[E_Pis_Name.V4020](
    sen_Open := gIO.i_EL[10].i_ch7,
    sen_Close := gIO.i_EL[10].i_ch8,
    DefaultCmd := E_PistonDefault_CMD.Close,
    iFB_Num := E_Pis_Name.V4020,
    stOperation := stOper[E_ModeZone.eCIP],
    valve_Open => GIO.q_Manifold2[3].sol_14); // FB_Piston

// NETWORK 27

// NETWORK 28
fbPis[E_Pis_Name.V4039](
    DefaultCmd := E_PistonDefault_CMD.Close,
    iFB_Num := E_Pis_Name.V4039,
    stOperation := stOper[E_ModeZone.eNone]); // FB_Piston

// NETWORK 29
fbPis[E_Pis_Name.V4040](
    sen_Open := gIO.i_EL[11].i_ch12,
    sen_Close := gIO.i_EL[11].i_ch11,
    DefaultCmd := E_PistonDefault_CMD.Open,
    iFB_Num := E_Pis_Name.V4040,
    stOperation := stOper[E_ModeZone.eTank4],
    valve_Close => GIO.q_Manifold2[10].sol_14); // FB_Piston

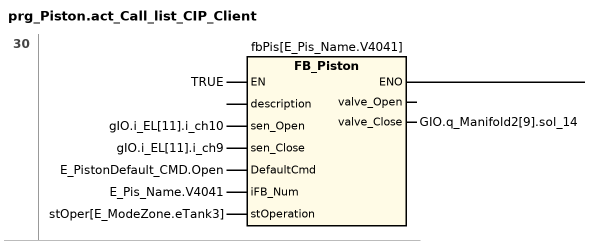
// NETWORK 30
fbPis[E_Pis_Name.V4041](
    sen_Open := gIO.i_EL[11].i_ch10,
    sen_Close := gIO.i_EL[11].i_ch9,
    DefaultCmd := E_PistonDefault_CMD.Open,
    iFB_Num := E_Pis_Name.V4041,
    stOperation := stOper[E_ModeZone.eTank3],
    valve_Close => GIO.q_Manifold2[9].sol_14); // FB_Piston
END_ACTION

ACTION act_Call_list_CIP_SourceNTarget:
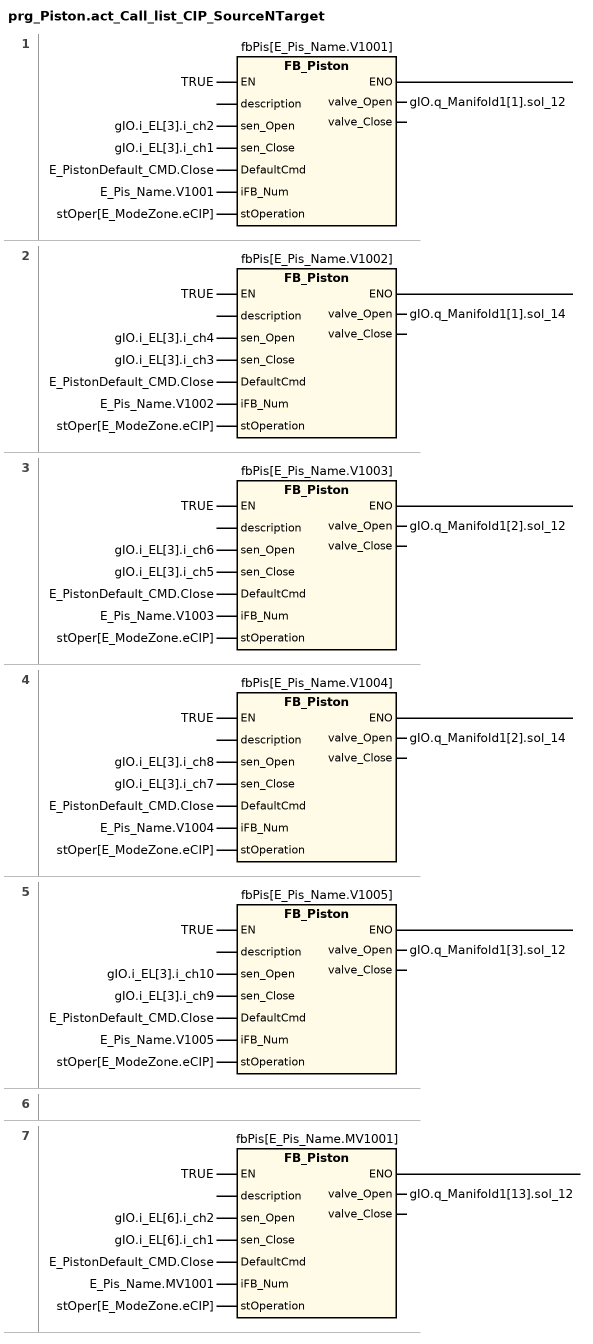
// NETWORK 1
fbPis[E_Pis_Name.V1001](
    sen_Open := gIO.i_EL[3].i_ch2,
    sen_Close := gIO.i_EL[3].i_ch1,
    DefaultCmd := E_PistonDefault_CMD.Close,
    iFB_Num := E_Pis_Name.V1001,
    stOperation := stOper[E_ModeZone.eCIP],
    valve_Open => gIO.q_Manifold1[1].sol_12); // FB_Piston

// NETWORK 2
fbPis[E_Pis_Name.V1002](
    sen_Open := gIO.i_EL[3].i_ch4,
    sen_Close := gIO.i_EL[3].i_ch3,
    DefaultCmd := E_PistonDefault_CMD.Close,
    iFB_Num := E_Pis_Name.V1002,
    stOperation := stOper[E_ModeZone.eCIP],
    valve_Open => gIO.q_Manifold1[1].sol_14); // FB_Piston

// NETWORK 3
fbPis[E_Pis_Name.V1003](
    sen_Open := gIO.i_EL[3].i_ch6,
    sen_Close := gIO.i_EL[3].i_ch5,
    DefaultCmd := E_PistonDefault_CMD.Close,
    iFB_Num := E_Pis_Name.V1003,
    stOperation := stOper[E_ModeZone.eCIP],
    valve_Open => gIO.q_Manifold1[2].sol_12); // FB_Piston

// NETWORK 4
fbPis[E_Pis_Name.V1004](
    sen_Open := gIO.i_EL[3].i_ch8,
    sen_Close := gIO.i_EL[3].i_ch7,
    DefaultCmd := E_PistonDefault_CMD.Close,
    iFB_Num := E_Pis_Name.V1004,
    stOperation := stOper[E_ModeZone.eCIP],
    valve_Open => gIO.q_Manifold1[2].sol_14); // FB_Piston

// NETWORK 5
fbPis[E_Pis_Name.V1005](
    sen_Open := gIO.i_EL[3].i_ch10,
    sen_Close := gIO.i_EL[3].i_ch9,
    DefaultCmd := E_PistonDefault_CMD.Close,
    iFB_Num := E_Pis_Name.V1005,
    stOperation := stOper[E_ModeZone.eCIP],
    valve_Open => gIO.q_Manifold1[3].sol_12); // FB_Piston

// NETWORK 6

// NETWORK 7
fbPis[E_Pis_Name.MV1001](
    sen_Open := gIO.i_EL[6].i_ch2,
    sen_Close := gIO.i_EL[6].i_ch1,
    DefaultCmd := E_PistonDefault_CMD.Close,
    iFB_Num := E_Pis_Name.MV1001,
    stOperation := stOper[E_ModeZone.eCIP],
    valve_Open => gIO.q_Manifold1[13].sol_12); // FB_Piston

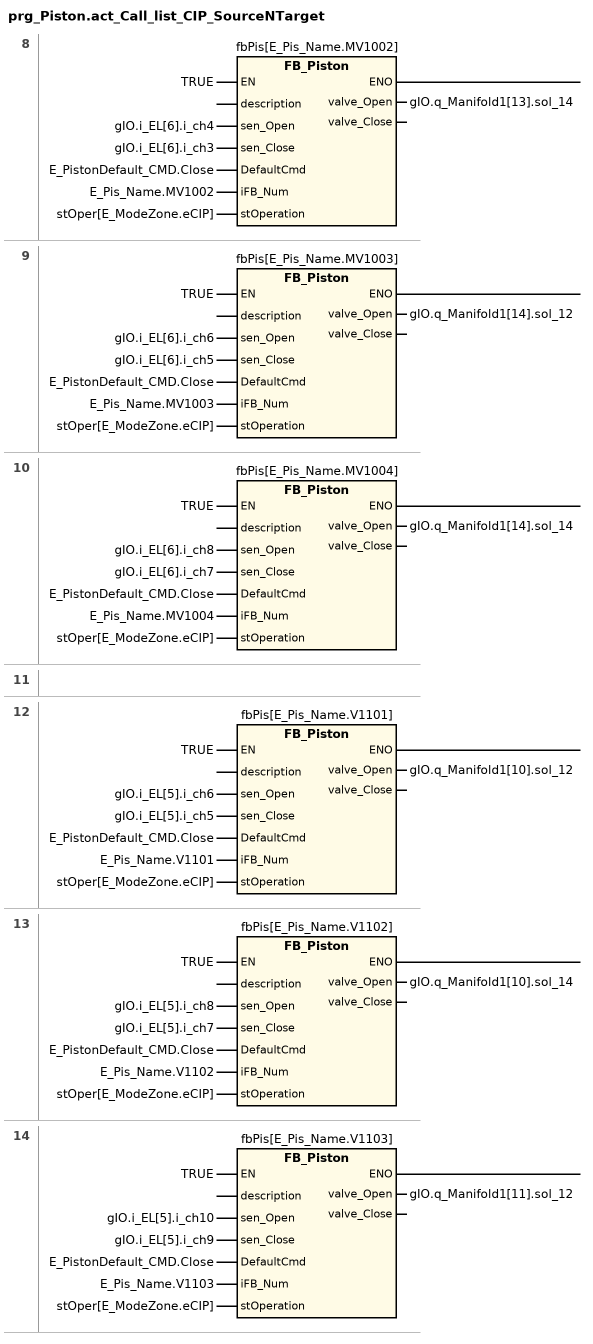
// NETWORK 8
fbPis[E_Pis_Name.MV1002](
    sen_Open := gIO.i_EL[6].i_ch4,
    sen_Close := gIO.i_EL[6].i_ch3,
    DefaultCmd := E_PistonDefault_CMD.Close,
    iFB_Num := E_Pis_Name.MV1002,
    stOperation := stOper[E_ModeZone.eCIP],
    valve_Open => gIO.q_Manifold1[13].sol_14); // FB_Piston

// NETWORK 9
fbPis[E_Pis_Name.MV1003](
    sen_Open := gIO.i_EL[6].i_ch6,
    sen_Close := gIO.i_EL[6].i_ch5,
    DefaultCmd := E_PistonDefault_CMD.Close,
    iFB_Num := E_Pis_Name.MV1003,
    stOperation := stOper[E_ModeZone.eCIP],
    valve_Open => gIO.q_Manifold1[14].sol_12); // FB_Piston

// NETWORK 10
fbPis[E_Pis_Name.MV1004](
    sen_Open := gIO.i_EL[6].i_ch8,
    sen_Close := gIO.i_EL[6].i_ch7,
    DefaultCmd := E_PistonDefault_CMD.Close,
    iFB_Num := E_Pis_Name.MV1004,
    stOperation := stOper[E_ModeZone.eCIP],
    valve_Open => gIO.q_Manifold1[14].sol_14); // FB_Piston

// NETWORK 11

// NETWORK 12
fbPis[E_Pis_Name.V1101](
    sen_Open := gIO.i_EL[5].i_ch6,
    sen_Close := gIO.i_EL[5].i_ch5,
    DefaultCmd := E_PistonDefault_CMD.Close,
    iFB_Num := E_Pis_Name.V1101,
    stOperation := stOper[E_ModeZone.eCIP],
    valve_Open => gIO.q_Manifold1[10].sol_12); // FB_Piston

// NETWORK 13
fbPis[E_Pis_Name.V1102](
    sen_Open := gIO.i_EL[5].i_ch8,
    sen_Close := gIO.i_EL[5].i_ch7,
    DefaultCmd := E_PistonDefault_CMD.Close,
    iFB_Num := E_Pis_Name.V1102,
    stOperation := stOper[E_ModeZone.eCIP],
    valve_Open => gIO.q_Manifold1[10].sol_14); // FB_Piston

// NETWORK 14
fbPis[E_Pis_Name.V1103](
    sen_Open := gIO.i_EL[5].i_ch10,
    sen_Close := gIO.i_EL[5].i_ch9,
    DefaultCmd := E_PistonDefault_CMD.Close,
    iFB_Num := E_Pis_Name.V1103,
    stOperation := stOper[E_ModeZone.eCIP],
    valve_Open => gIO.q_Manifold1[11].sol_12); // FB_Piston

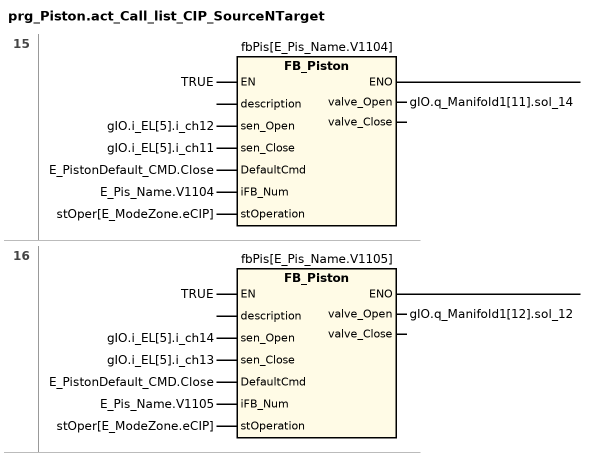
// NETWORK 15
fbPis[E_Pis_Name.V1104](
    sen_Open := gIO.i_EL[5].i_ch12,
    sen_Close := gIO.i_EL[5].i_ch11,
    DefaultCmd := E_PistonDefault_CMD.Close,
    iFB_Num := E_Pis_Name.V1104,
    stOperation := stOper[E_ModeZone.eCIP],
    valve_Open => gIO.q_Manifold1[11].sol_14); // FB_Piston

// NETWORK 16
fbPis[E_Pis_Name.V1105](
    sen_Open := gIO.i_EL[5].i_ch14,
    sen_Close := gIO.i_EL[5].i_ch13,
    DefaultCmd := E_PistonDefault_CMD.Close,
    iFB_Num := E_Pis_Name.V1105,
    stOperation := stOper[E_ModeZone.eCIP],
    valve_Open => gIO.q_Manifold1[12].sol_12); // FB_Piston
END_ACTION

ACTION act_Call_list_CIP_Tanks:
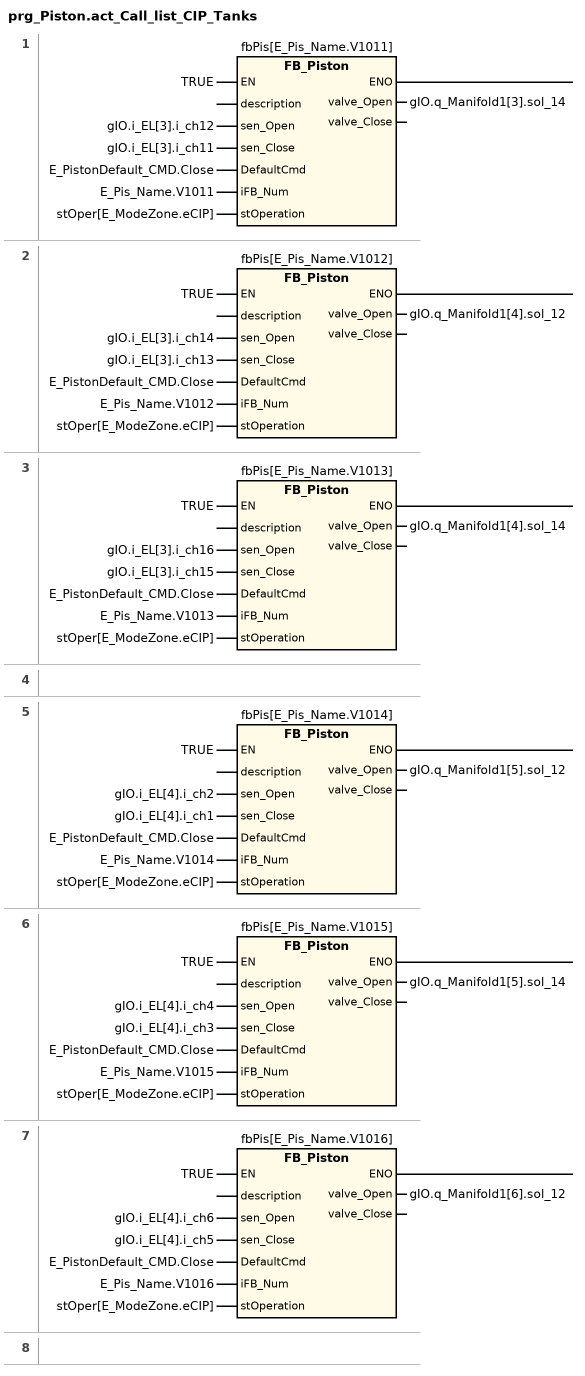
// NETWORK 1
fbPis[E_Pis_Name.V1011](
    sen_Open := gIO.i_EL[3].i_ch12,
    sen_Close := gIO.i_EL[3].i_ch11,
    DefaultCmd := E_PistonDefault_CMD.Close,
    iFB_Num := E_Pis_Name.V1011,
    stOperation := stOper[E_ModeZone.eCIP],
    valve_Open => gIO.q_Manifold1[3].sol_14); // FB_Piston

// NETWORK 2
fbPis[E_Pis_Name.V1012](
    sen_Open := gIO.i_EL[3].i_ch14,
    sen_Close := gIO.i_EL[3].i_ch13,
    DefaultCmd := E_PistonDefault_CMD.Close,
    iFB_Num := E_Pis_Name.V1012,
    stOperation := stOper[E_ModeZone.eCIP],
    valve_Open => gIO.q_Manifold1[4].sol_12); // FB_Piston

// NETWORK 3
fbPis[E_Pis_Name.V1013](
    sen_Open := gIO.i_EL[3].i_ch16,
    sen_Close := gIO.i_EL[3].i_ch15,
    DefaultCmd := E_PistonDefault_CMD.Close,
    iFB_Num := E_Pis_Name.V1013,
    stOperation := stOper[E_ModeZone.eCIP],
    valve_Open => gIO.q_Manifold1[4].sol_14); // FB_Piston

// NETWORK 4

// NETWORK 5
fbPis[E_Pis_Name.V1014](
    sen_Open := gIO.i_EL[4].i_ch2,
    sen_Close := gIO.i_EL[4].i_ch1,
    DefaultCmd := E_PistonDefault_CMD.Close,
    iFB_Num := E_Pis_Name.V1014,
    stOperation := stOper[E_ModeZone.eCIP],
    valve_Open => gIO.q_Manifold1[5].sol_12); // FB_Piston

// NETWORK 6
fbPis[E_Pis_Name.V1015](
    sen_Open := gIO.i_EL[4].i_ch4,
    sen_Close := gIO.i_EL[4].i_ch3,
    DefaultCmd := E_PistonDefault_CMD.Close,
    iFB_Num := E_Pis_Name.V1015,
    stOperation := stOper[E_ModeZone.eCIP],
    valve_Open => gIO.q_Manifold1[5].sol_14); // FB_Piston

// NETWORK 7
fbPis[E_Pis_Name.V1016](
    sen_Open := gIO.i_EL[4].i_ch6,
    sen_Close := gIO.i_EL[4].i_ch5,
    DefaultCmd := E_PistonDefault_CMD.Close,
    iFB_Num := E_Pis_Name.V1016,
    stOperation := stOper[E_ModeZone.eCIP],
    valve_Open => gIO.q_Manifold1[6].sol_12); // FB_Piston

// NETWORK 8

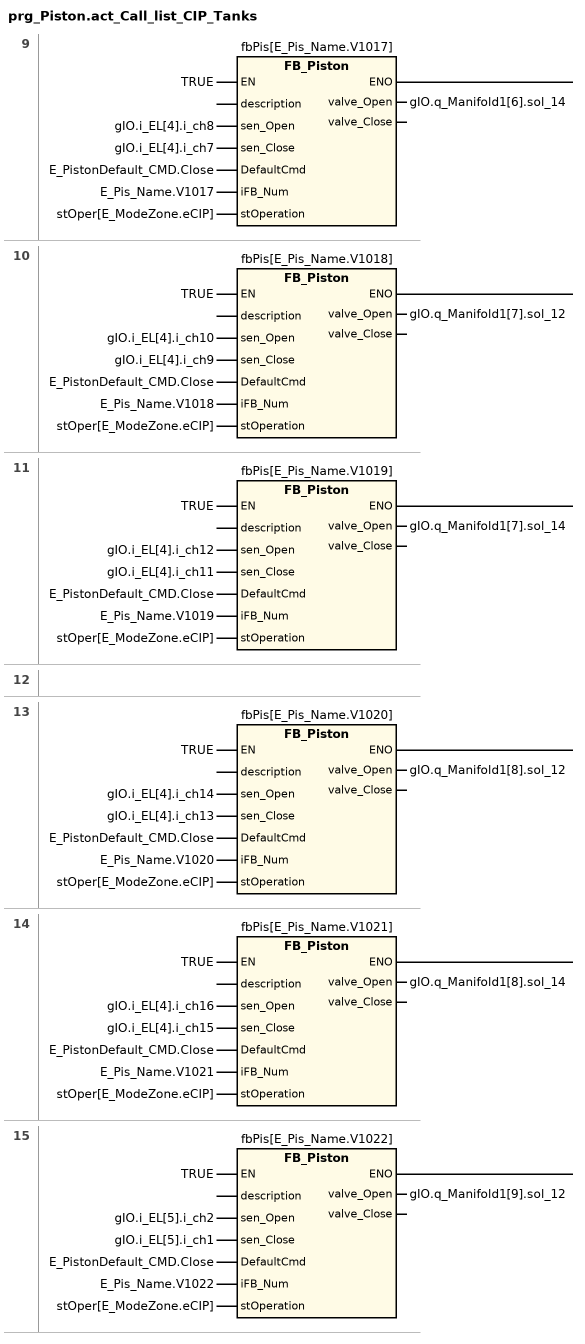
// NETWORK 9
fbPis[E_Pis_Name.V1017](
    sen_Open := gIO.i_EL[4].i_ch8,
    sen_Close := gIO.i_EL[4].i_ch7,
    DefaultCmd := E_PistonDefault_CMD.Close,
    iFB_Num := E_Pis_Name.V1017,
    stOperation := stOper[E_ModeZone.eCIP],
    valve_Open => gIO.q_Manifold1[6].sol_14); // FB_Piston

// NETWORK 10
fbPis[E_Pis_Name.V1018](
    sen_Open := gIO.i_EL[4].i_ch10,
    sen_Close := gIO.i_EL[4].i_ch9,
    DefaultCmd := E_PistonDefault_CMD.Close,
    iFB_Num := E_Pis_Name.V1018,
    stOperation := stOper[E_ModeZone.eCIP],
    valve_Open => gIO.q_Manifold1[7].sol_12); // FB_Piston

// NETWORK 11
fbPis[E_Pis_Name.V1019](
    sen_Open := gIO.i_EL[4].i_ch12,
    sen_Close := gIO.i_EL[4].i_ch11,
    DefaultCmd := E_PistonDefault_CMD.Close,
    iFB_Num := E_Pis_Name.V1019,
    stOperation := stOper[E_ModeZone.eCIP],
    valve_Open => gIO.q_Manifold1[7].sol_14); // FB_Piston

// NETWORK 12

// NETWORK 13
fbPis[E_Pis_Name.V1020](
    sen_Open := gIO.i_EL[4].i_ch14,
    sen_Close := gIO.i_EL[4].i_ch13,
    DefaultCmd := E_PistonDefault_CMD.Close,
    iFB_Num := E_Pis_Name.V1020,
    stOperation := stOper[E_ModeZone.eCIP],
    valve_Open => gIO.q_Manifold1[8].sol_12); // FB_Piston

// NETWORK 14
fbPis[E_Pis_Name.V1021](
    sen_Open := gIO.i_EL[4].i_ch16,
    sen_Close := gIO.i_EL[4].i_ch15,
    DefaultCmd := E_PistonDefault_CMD.Close,
    iFB_Num := E_Pis_Name.V1021,
    stOperation := stOper[E_ModeZone.eCIP],
    valve_Open => gIO.q_Manifold1[8].sol_14); // FB_Piston

// NETWORK 15
fbPis[E_Pis_Name.V1022](
    sen_Open := gIO.i_EL[5].i_ch2,
    sen_Close := gIO.i_EL[5].i_ch1,
    DefaultCmd := E_PistonDefault_CMD.Close,
    iFB_Num := E_Pis_Name.V1022,
    stOperation := stOper[E_ModeZone.eCIP],
    valve_Open => gIO.q_Manifold1[9].sol_12); // FB_Piston

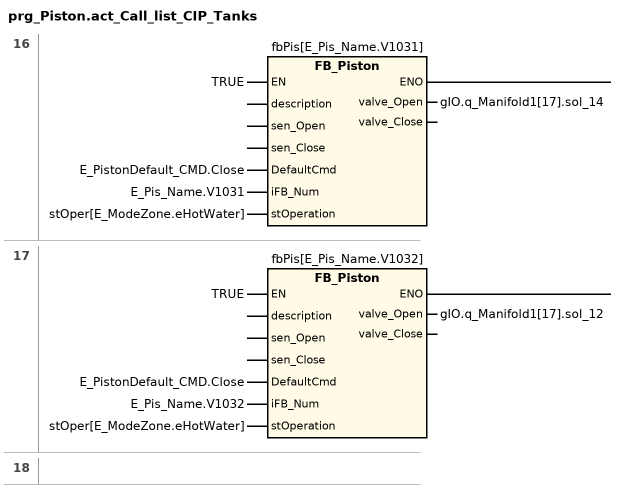
// NETWORK 16
fbPis[E_Pis_Name.V1031](
    DefaultCmd := E_PistonDefault_CMD.Close,
    iFB_Num := E_Pis_Name.V1031,
    stOperation := stOper[E_ModeZone.eHotWater],
    valve_Open => gIO.q_Manifold1[17].sol_14); // FB_Piston

// NETWORK 17
fbPis[E_Pis_Name.V1032](
    DefaultCmd := E_PistonDefault_CMD.Close,
    iFB_Num := E_Pis_Name.V1032,
    stOperation := stOper[E_ModeZone.eHotWater],
    valve_Open => gIO.q_Manifold1[17].sol_12); // FB_Piston

// NETWORK 18
END_ACTION

ACTION act_Call_List_LineSource:
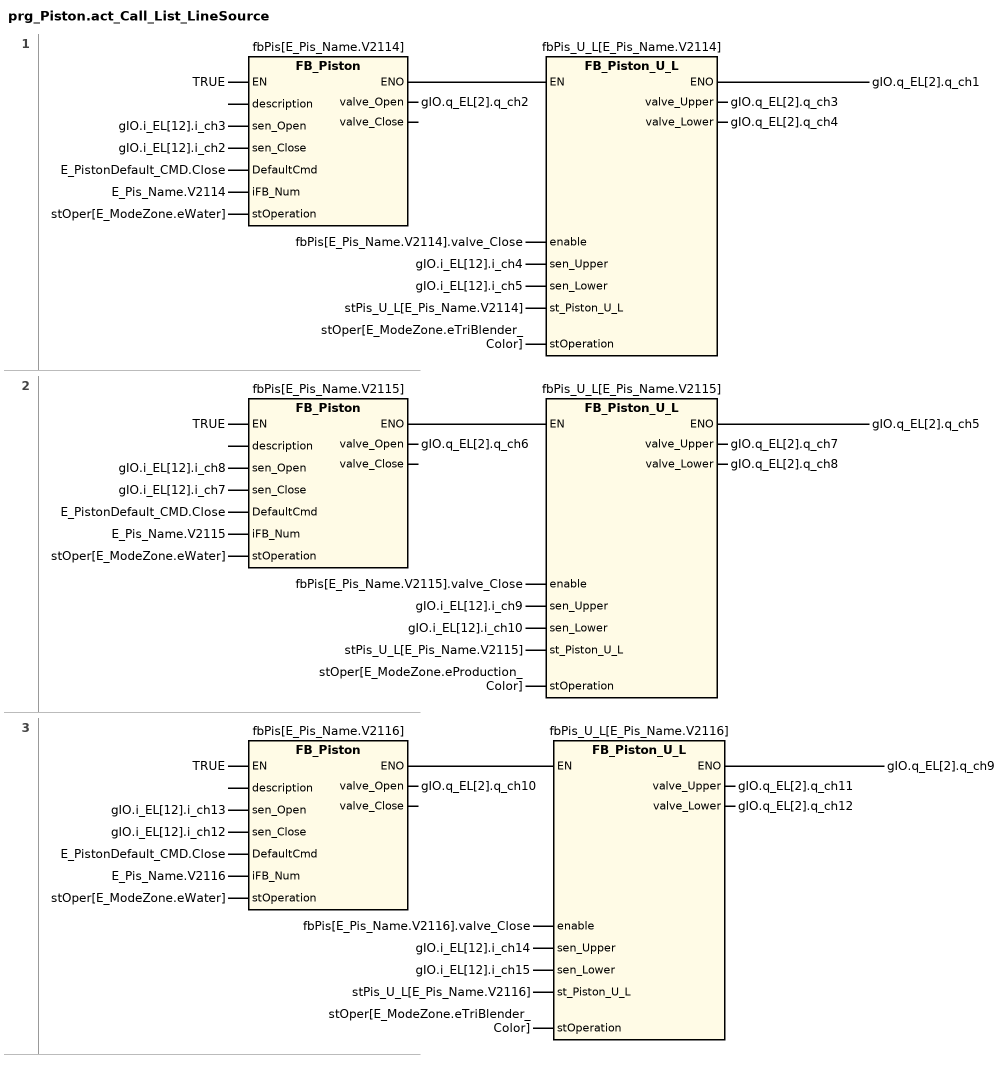
// NETWORK 1
fbPis[E_Pis_Name.V2114](
    sen_Open := gIO.i_EL[12].i_ch3,
    sen_Close := gIO.i_EL[12].i_ch2,
    DefaultCmd := E_PistonDefault_CMD.Close,
    iFB_Num := E_Pis_Name.V2114,
    stOperation := stOper[E_ModeZone.eWater],
    valve_Open => gIO.q_EL[2].q_ch2); // FB_Piston
fbPis_U_L[E_Pis_Name.V2114](
    enable := fbPis[E_Pis_Name.V2114].valve_Close,
    sen_Upper := gIO.i_EL[12].i_ch4,
    sen_Lower := gIO.i_EL[12].i_ch5,
    st_Piston_U_L := stPis_U_L[E_Pis_Name.V2114],
    stOperation := stOper[E_ModeZone.eTriBlender_Color],
    valve_Upper => gIO.q_EL[2].q_ch3,
    valve_Lower => gIO.q_EL[2].q_ch4); // FB_Piston_U_L
gIO.q_EL[2].q_ch1 := TRUE;

// NETWORK 2
fbPis[E_Pis_Name.V2115](
    sen_Open := gIO.i_EL[12].i_ch8,
    sen_Close := gIO.i_EL[12].i_ch7,
    DefaultCmd := E_PistonDefault_CMD.Close,
    iFB_Num := E_Pis_Name.V2115,
    stOperation := stOper[E_ModeZone.eWater],
    valve_Open => gIO.q_EL[2].q_ch6); // FB_Piston
fbPis_U_L[E_Pis_Name.V2115](
    enable := fbPis[E_Pis_Name.V2115].valve_Close,
    sen_Upper := gIO.i_EL[12].i_ch9,
    sen_Lower := gIO.i_EL[12].i_ch10,
    st_Piston_U_L := stPis_U_L[E_Pis_Name.V2115],
    stOperation := stOper[E_ModeZone.eProduction_Color],
    valve_Upper => gIO.q_EL[2].q_ch7,
    valve_Lower => gIO.q_EL[2].q_ch8); // FB_Piston_U_L
gIO.q_EL[2].q_ch5 := TRUE;

// NETWORK 3
fbPis[E_Pis_Name.V2116](
    sen_Open := gIO.i_EL[12].i_ch13,
    sen_Close := gIO.i_EL[12].i_ch12,
    DefaultCmd := E_PistonDefault_CMD.Close,
    iFB_Num := E_Pis_Name.V2116,
    stOperation := stOper[E_ModeZone.eWater],
    valve_Open => gIO.q_EL[2].q_ch10); // FB_Piston
fbPis_U_L[E_Pis_Name.V2116](
    enable := fbPis[E_Pis_Name.V2116].valve_Close,
    sen_Upper := gIO.i_EL[12].i_ch14,
    sen_Lower := gIO.i_EL[12].i_ch15,
    st_Piston_U_L := stPis_U_L[E_Pis_Name.V2116],
    stOperation := stOper[E_ModeZone.eTriBlender_Color],
    valve_Upper => gIO.q_EL[2].q_ch11,
    valve_Lower => gIO.q_EL[2].q_ch12); // FB_Piston_U_L
gIO.q_EL[2].q_ch9 := TRUE;

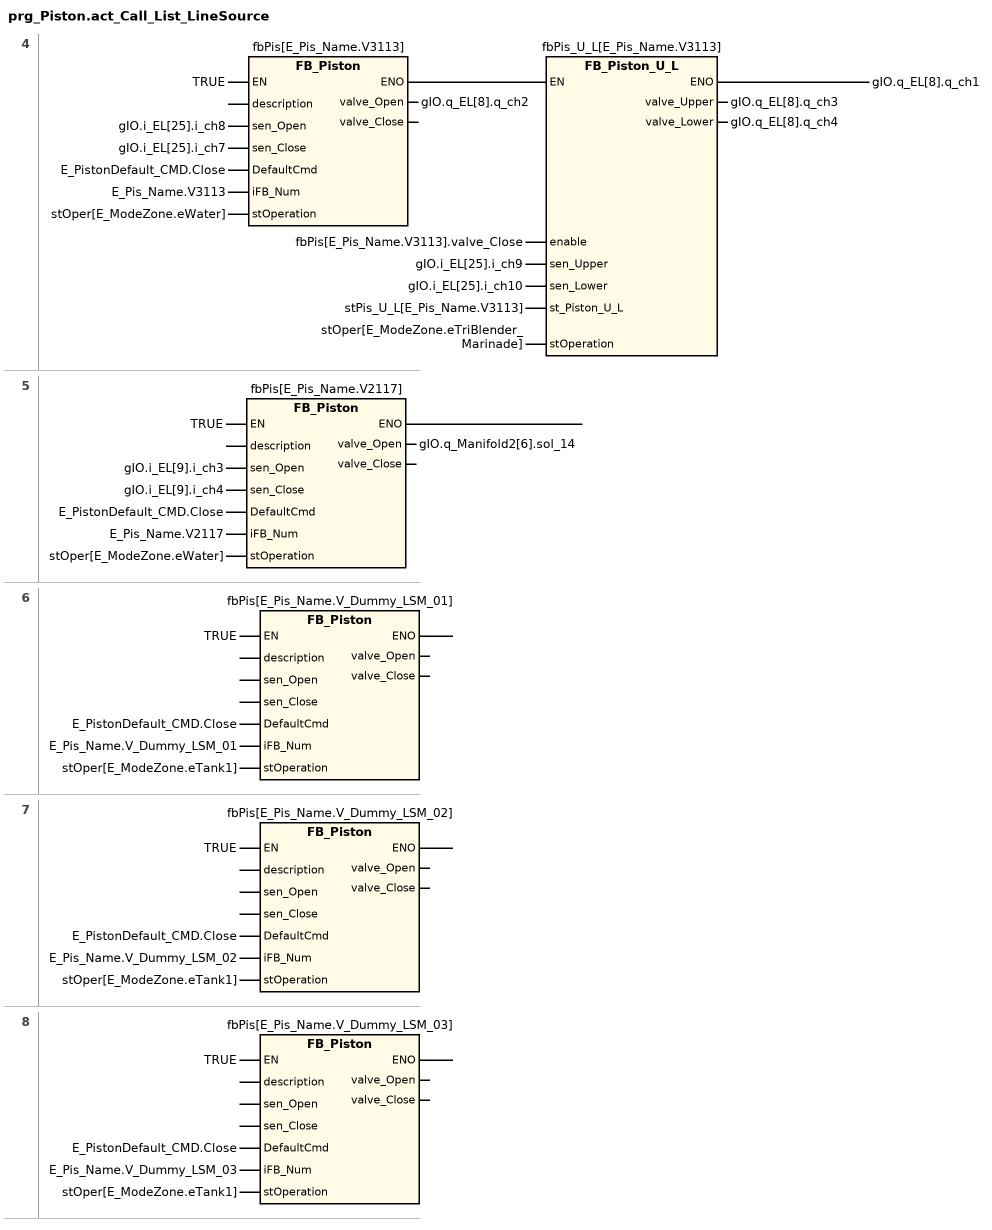
// NETWORK 4
fbPis[E_Pis_Name.V3113](
    sen_Open := gIO.i_EL[25].i_ch8,
    sen_Close := gIO.i_EL[25].i_ch7,
    DefaultCmd := E_PistonDefault_CMD.Close,
    iFB_Num := E_Pis_Name.V3113,
    stOperation := stOper[E_ModeZone.eWater],
    valve_Open => gIO.q_EL[8].q_ch2); // FB_Piston
fbPis_U_L[E_Pis_Name.V3113](
    enable := fbPis[E_Pis_Name.V3113].valve_Close,
    sen_Upper := gIO.i_EL[25].i_ch9,
    sen_Lower := gIO.i_EL[25].i_ch10,
    st_Piston_U_L := stPis_U_L[E_Pis_Name.V3113],
    stOperation := stOper[E_ModeZone.eTriBlender_Marinade],
    valve_Upper => gIO.q_EL[8].q_ch3,
    valve_Lower => gIO.q_EL[8].q_ch4); // FB_Piston_U_L
gIO.q_EL[8].q_ch1 := TRUE;

// NETWORK 5
fbPis[E_Pis_Name.V2117](
    sen_Open := gIO.i_EL[9].i_ch3,
    sen_Close := gIO.i_EL[9].i_ch4,
    DefaultCmd := E_PistonDefault_CMD.Close,
    iFB_Num := E_Pis_Name.V2117,
    stOperation := stOper[E_ModeZone.eWater],
    valve_Open => gIO.q_Manifold2[6].sol_14); // FB_Piston

// NETWORK 6
fbPis[E_Pis_Name.V_Dummy_LSM_01](
    DefaultCmd := E_PistonDefault_CMD.Close,
    iFB_Num := E_Pis_Name.V_Dummy_LSM_01,
    stOperation := stOper[E_ModeZone.eTank1]); // FB_Piston

// NETWORK 7
fbPis[E_Pis_Name.V_Dummy_LSM_02](
    DefaultCmd := E_PistonDefault_CMD.Close,
    iFB_Num := E_Pis_Name.V_Dummy_LSM_02,
    stOperation := stOper[E_ModeZone.eTank1]); // FB_Piston

// NETWORK 8
fbPis[E_Pis_Name.V_Dummy_LSM_03](
    DefaultCmd := E_PistonDefault_CMD.Close,
    iFB_Num := E_Pis_Name.V_Dummy_LSM_03,
    stOperation := stOper[E_ModeZone.eTank1]); // FB_Piston

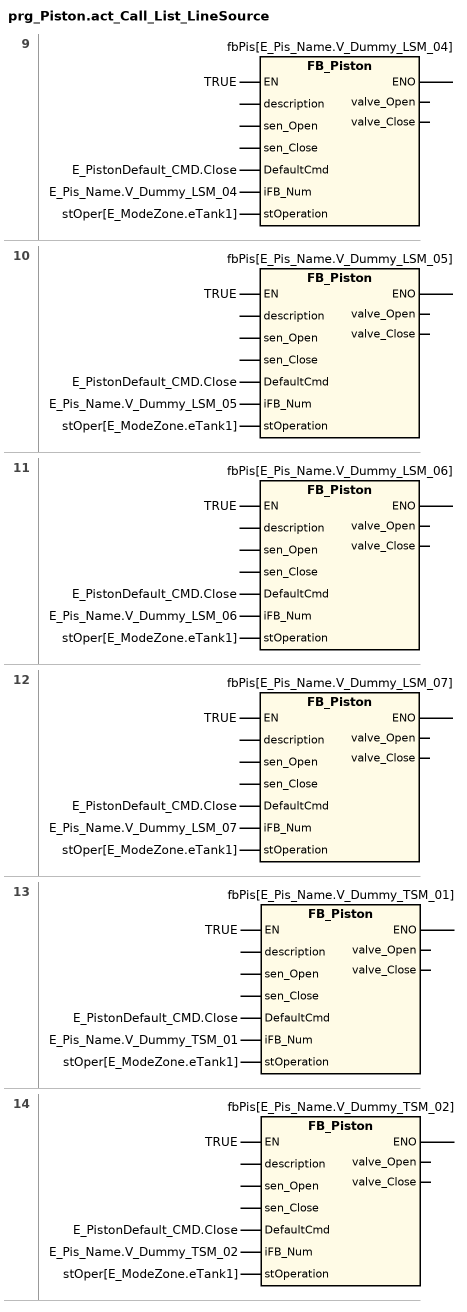
// NETWORK 9
fbPis[E_Pis_Name.V_Dummy_LSM_04](
    DefaultCmd := E_PistonDefault_CMD.Close,
    iFB_Num := E_Pis_Name.V_Dummy_LSM_04,
    stOperation := stOper[E_ModeZone.eTank1]); // FB_Piston

// NETWORK 10
fbPis[E_Pis_Name.V_Dummy_LSM_05](
    DefaultCmd := E_PistonDefault_CMD.Close,
    iFB_Num := E_Pis_Name.V_Dummy_LSM_05,
    stOperation := stOper[E_ModeZone.eTank1]); // FB_Piston

// NETWORK 11
fbPis[E_Pis_Name.V_Dummy_LSM_06](
    DefaultCmd := E_PistonDefault_CMD.Close,
    iFB_Num := E_Pis_Name.V_Dummy_LSM_06,
    stOperation := stOper[E_ModeZone.eTank1]); // FB_Piston

// NETWORK 12
fbPis[E_Pis_Name.V_Dummy_LSM_07](
    DefaultCmd := E_PistonDefault_CMD.Close,
    iFB_Num := E_Pis_Name.V_Dummy_LSM_07,
    stOperation := stOper[E_ModeZone.eTank1]); // FB_Piston

// NETWORK 13
fbPis[E_Pis_Name.V_Dummy_TSM_01](
    DefaultCmd := E_PistonDefault_CMD.Close,
    iFB_Num := E_Pis_Name.V_Dummy_TSM_01,
    stOperation := stOper[E_ModeZone.eTank1]); // FB_Piston

// NETWORK 14
fbPis[E_Pis_Name.V_Dummy_TSM_02](
    DefaultCmd := E_PistonDefault_CMD.Close,
    iFB_Num := E_Pis_Name.V_Dummy_TSM_02,
    stOperation := stOper[E_ModeZone.eTank1]); // FB_Piston

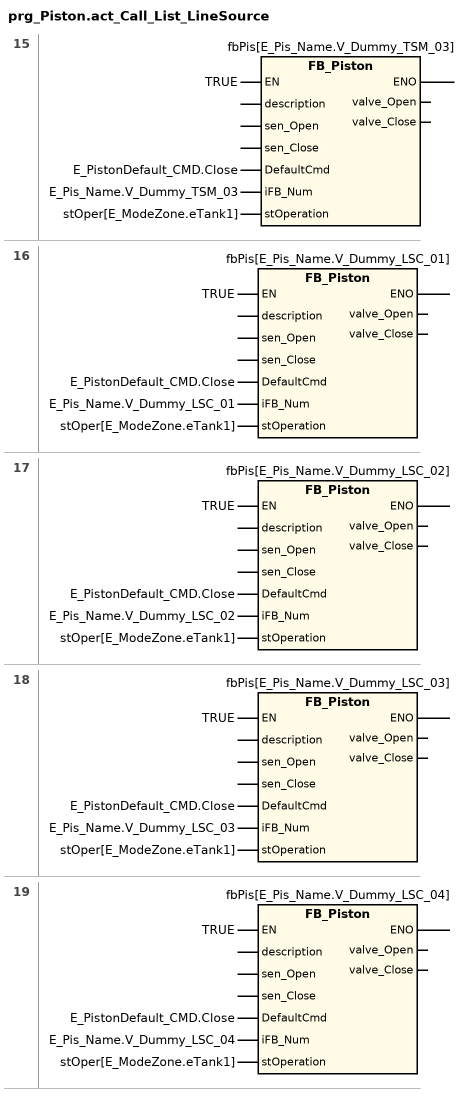
// NETWORK 15
fbPis[E_Pis_Name.V_Dummy_TSM_03](
    DefaultCmd := E_PistonDefault_CMD.Close,
    iFB_Num := E_Pis_Name.V_Dummy_TSM_03,
    stOperation := stOper[E_ModeZone.eTank1]); // FB_Piston

// NETWORK 16
fbPis[E_Pis_Name.V_Dummy_LSC_01](
    DefaultCmd := E_PistonDefault_CMD.Close,
    iFB_Num := E_Pis_Name.V_Dummy_LSC_01,
    stOperation := stOper[E_ModeZone.eTank1]); // FB_Piston

// NETWORK 17
fbPis[E_Pis_Name.V_Dummy_LSC_02](
    DefaultCmd := E_PistonDefault_CMD.Close,
    iFB_Num := E_Pis_Name.V_Dummy_LSC_02,
    stOperation := stOper[E_ModeZone.eTank1]); // FB_Piston

// NETWORK 18
fbPis[E_Pis_Name.V_Dummy_LSC_03](
    DefaultCmd := E_PistonDefault_CMD.Close,
    iFB_Num := E_Pis_Name.V_Dummy_LSC_03,
    stOperation := stOper[E_ModeZone.eTank1]); // FB_Piston

// NETWORK 19
fbPis[E_Pis_Name.V_Dummy_LSC_04](
    DefaultCmd := E_PistonDefault_CMD.Close,
    iFB_Num := E_Pis_Name.V_Dummy_LSC_04,
    stOperation := stOper[E_ModeZone.eTank1]); // FB_Piston
END_ACTION

ACTION act_Call_List_LineTarget:
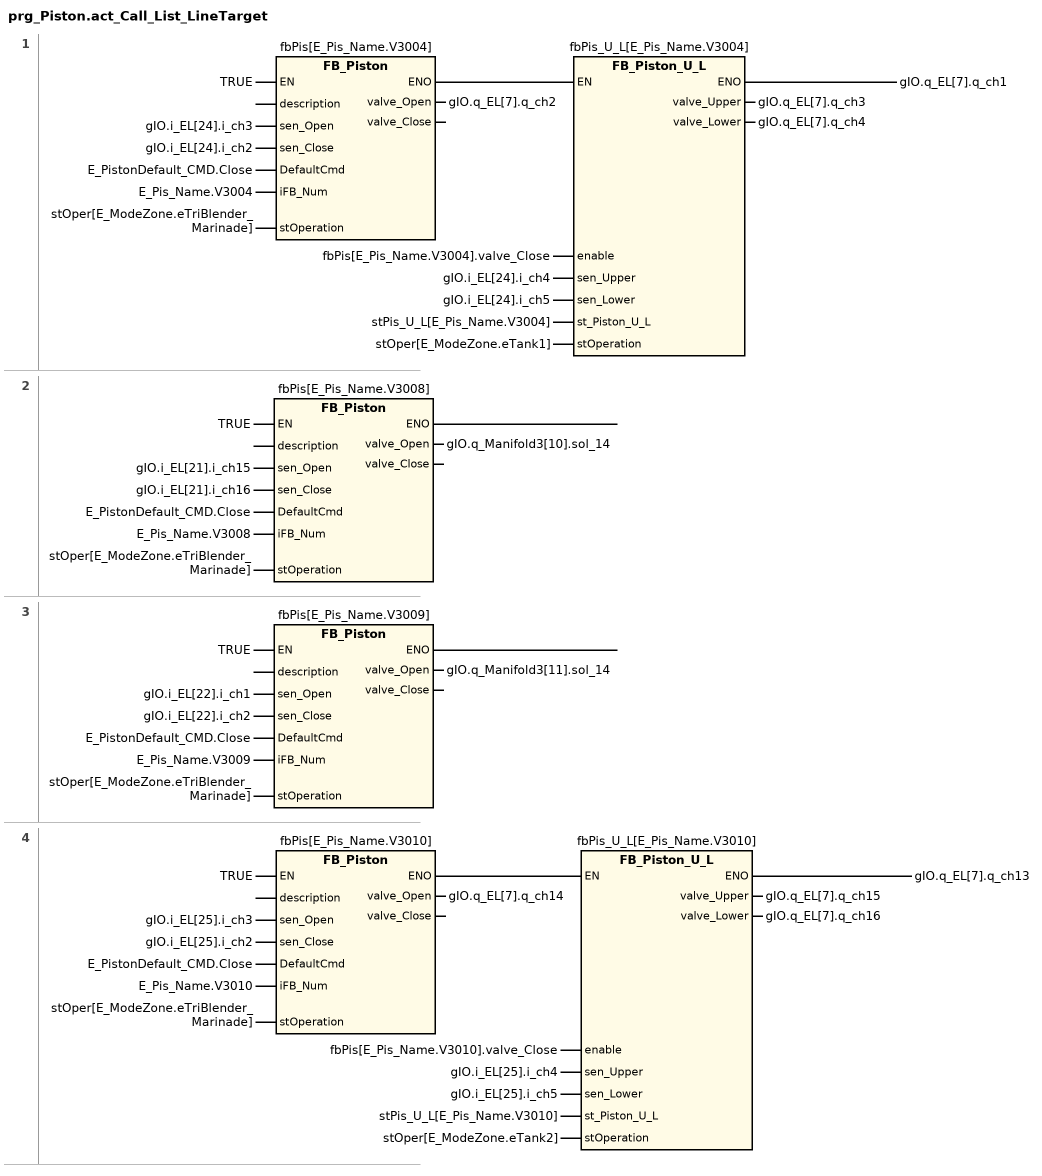
// NETWORK 1
fbPis[E_Pis_Name.V3004](
    sen_Open := gIO.i_EL[24].i_ch3,
    sen_Close := gIO.i_EL[24].i_ch2,
    DefaultCmd := E_PistonDefault_CMD.Close,
    iFB_Num := E_Pis_Name.V3004,
    stOperation := stOper[E_ModeZone.eTriBlender_Marinade],
    valve_Open => gIO.q_EL[7].q_ch2); // FB_Piston
fbPis_U_L[E_Pis_Name.V3004](
    enable := fbPis[E_Pis_Name.V3004].valve_Close,
    sen_Upper := gIO.i_EL[24].i_ch4,
    sen_Lower := gIO.i_EL[24].i_ch5,
    st_Piston_U_L := stPis_U_L[E_Pis_Name.V3004],
    stOperation := stOper[E_ModeZone.eTank1],
    valve_Upper => gIO.q_EL[7].q_ch3,
    valve_Lower => gIO.q_EL[7].q_ch4); // FB_Piston_U_L
gIO.q_EL[7].q_ch1 := TRUE;

// NETWORK 2
fbPis[E_Pis_Name.V3008](
    sen_Open := gIO.i_EL[21].i_ch15,
    sen_Close := gIO.i_EL[21].i_ch16,
    DefaultCmd := E_PistonDefault_CMD.Close,
    iFB_Num := E_Pis_Name.V3008,
    stOperation := stOper[E_ModeZone.eTriBlender_Marinade],
    valve_Open => gIO.q_Manifold3[10].sol_14); // FB_Piston

// NETWORK 3
fbPis[E_Pis_Name.V3009](
    sen_Open := gIO.i_EL[22].i_ch1,
    sen_Close := gIO.i_EL[22].i_ch2,
    DefaultCmd := E_PistonDefault_CMD.Close,
    iFB_Num := E_Pis_Name.V3009,
    stOperation := stOper[E_ModeZone.eTriBlender_Marinade],
    valve_Open => gIO.q_Manifold3[11].sol_14); // FB_Piston

// NETWORK 4
fbPis[E_Pis_Name.V3010](
    sen_Open := gIO.i_EL[25].i_ch3,
    sen_Close := gIO.i_EL[25].i_ch2,
    DefaultCmd := E_PistonDefault_CMD.Close,
    iFB_Num := E_Pis_Name.V3010,
    stOperation := stOper[E_ModeZone.eTriBlender_Marinade],
    valve_Open => gIO.q_EL[7].q_ch14); // FB_Piston
fbPis_U_L[E_Pis_Name.V3010](
    enable := fbPis[E_Pis_Name.V3010].valve_Close,
    sen_Upper := gIO.i_EL[25].i_ch4,
    sen_Lower := gIO.i_EL[25].i_ch5,
    st_Piston_U_L := stPis_U_L[E_Pis_Name.V3010],
    stOperation := stOper[E_ModeZone.eTank2],
    valve_Upper => gIO.q_EL[7].q_ch15,
    valve_Lower => gIO.q_EL[7].q_ch16); // FB_Piston_U_L
gIO.q_EL[7].q_ch13 := TRUE;

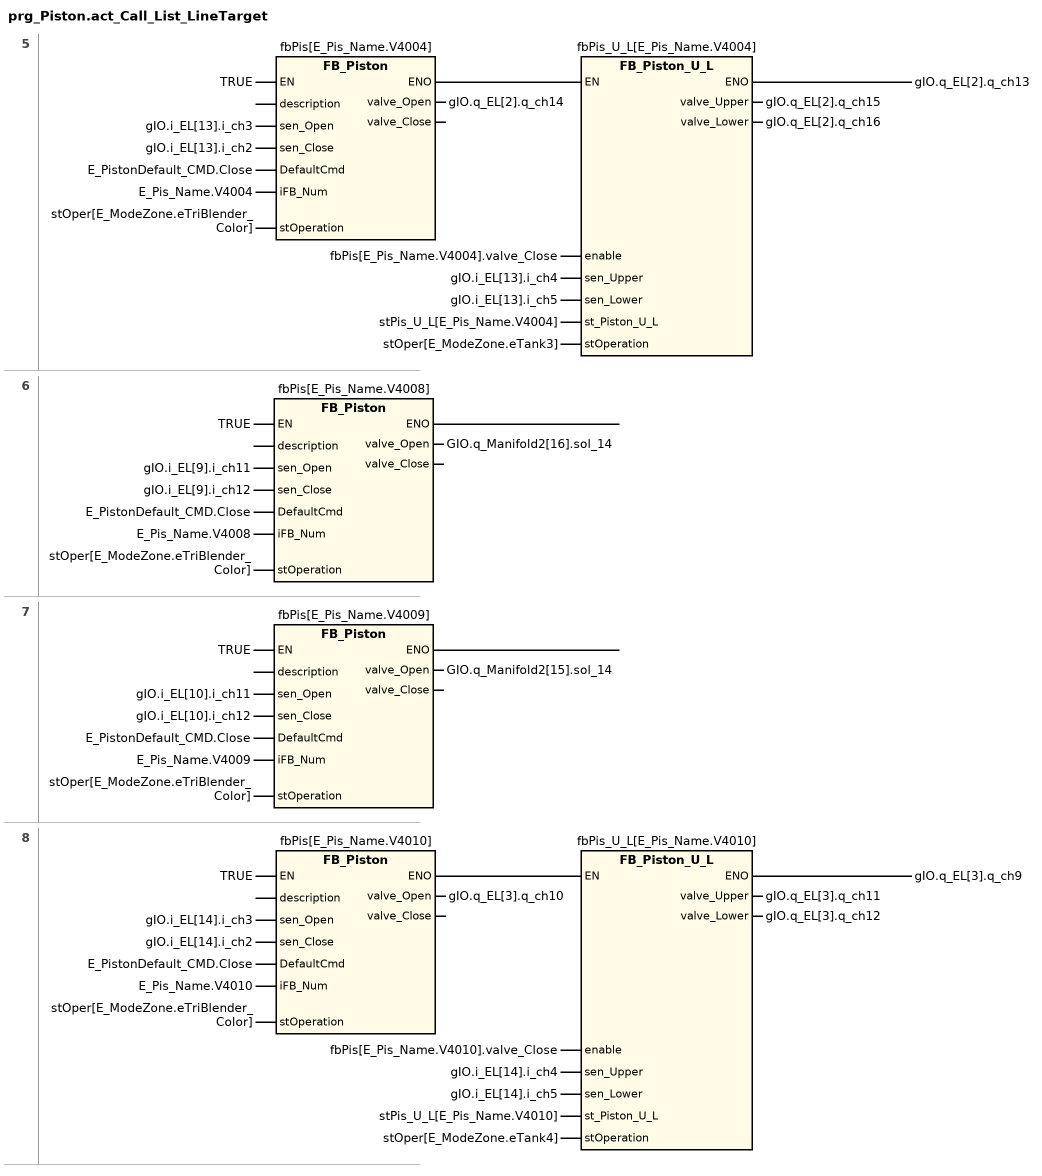
// NETWORK 5
fbPis[E_Pis_Name.V4004](
    sen_Open := gIO.i_EL[13].i_ch3,
    sen_Close := gIO.i_EL[13].i_ch2,
    DefaultCmd := E_PistonDefault_CMD.Close,
    iFB_Num := E_Pis_Name.V4004,
    stOperation := stOper[E_ModeZone.eTriBlender_Color],
    valve_Open => gIO.q_EL[2].q_ch14); // FB_Piston
fbPis_U_L[E_Pis_Name.V4004](
    enable := fbPis[E_Pis_Name.V4004].valve_Close,
    sen_Upper := gIO.i_EL[13].i_ch4,
    sen_Lower := gIO.i_EL[13].i_ch5,
    st_Piston_U_L := stPis_U_L[E_Pis_Name.V4004],
    stOperation := stOper[E_ModeZone.eTank3],
    valve_Upper => gIO.q_EL[2].q_ch15,
    valve_Lower => gIO.q_EL[2].q_ch16); // FB_Piston_U_L
gIO.q_EL[2].q_ch13 := TRUE;

// NETWORK 6
fbPis[E_Pis_Name.V4008](
    sen_Open := gIO.i_EL[9].i_ch11,
    sen_Close := gIO.i_EL[9].i_ch12,
    DefaultCmd := E_PistonDefault_CMD.Close,
    iFB_Num := E_Pis_Name.V4008,
    stOperation := stOper[E_ModeZone.eTriBlender_Color],
    valve_Open => GIO.q_Manifold2[16].sol_14); // FB_Piston

// NETWORK 7
fbPis[E_Pis_Name.V4009](
    sen_Open := gIO.i_EL[10].i_ch11,
    sen_Close := gIO.i_EL[10].i_ch12,
    DefaultCmd := E_PistonDefault_CMD.Close,
    iFB_Num := E_Pis_Name.V4009,
    stOperation := stOper[E_ModeZone.eTriBlender_Color],
    valve_Open => GIO.q_Manifold2[15].sol_14); // FB_Piston

// NETWORK 8
fbPis[E_Pis_Name.V4010](
    sen_Open := gIO.i_EL[14].i_ch3,
    sen_Close := gIO.i_EL[14].i_ch2,
    DefaultCmd := E_PistonDefault_CMD.Close,
    iFB_Num := E_Pis_Name.V4010,
    stOperation := stOper[E_ModeZone.eTriBlender_Color],
    valve_Open => gIO.q_EL[3].q_ch10); // FB_Piston
fbPis_U_L[E_Pis_Name.V4010](
    enable := fbPis[E_Pis_Name.V4010].valve_Close,
    sen_Upper := gIO.i_EL[14].i_ch4,
    sen_Lower := gIO.i_EL[14].i_ch5,
    st_Piston_U_L := stPis_U_L[E_Pis_Name.V4010],
    stOperation := stOper[E_ModeZone.eTank4],
    valve_Upper => gIO.q_EL[3].q_ch11,
    valve_Lower => gIO.q_EL[3].q_ch12); // FB_Piston_U_L
gIO.q_EL[3].q_ch9 := TRUE;

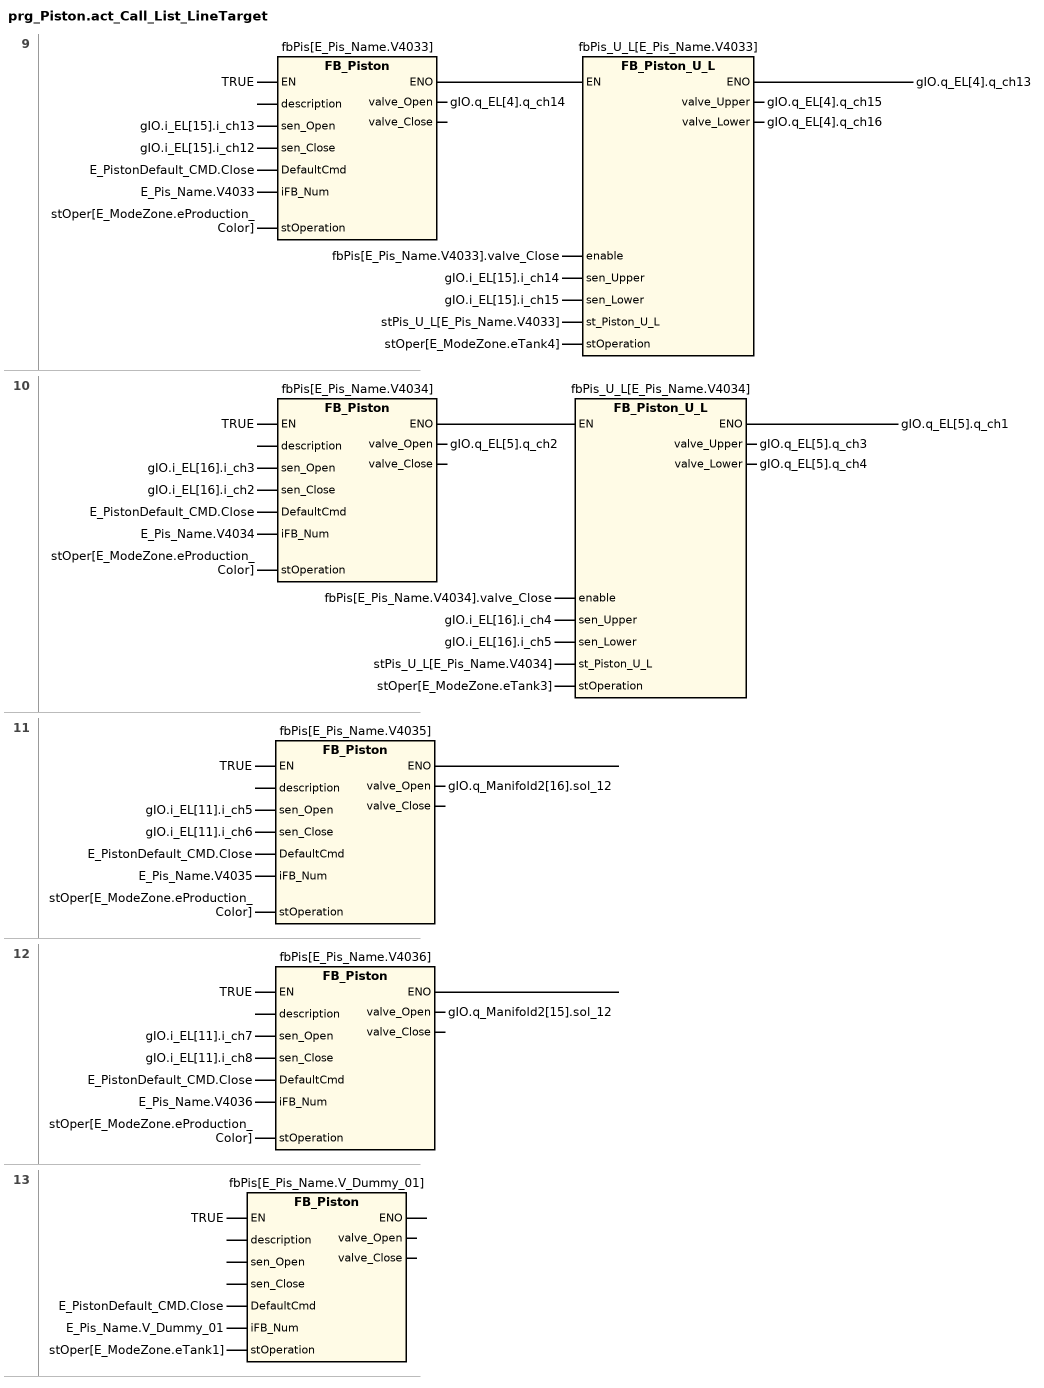
// NETWORK 9
fbPis[E_Pis_Name.V4033](
    sen_Open := gIO.i_EL[15].i_ch13,
    sen_Close := gIO.i_EL[15].i_ch12,
    DefaultCmd := E_PistonDefault_CMD.Close,
    iFB_Num := E_Pis_Name.V4033,
    stOperation := stOper[E_ModeZone.eProduction_Color],
    valve_Open => gIO.q_EL[4].q_ch14); // FB_Piston
fbPis_U_L[E_Pis_Name.V4033](
    enable := fbPis[E_Pis_Name.V4033].valve_Close,
    sen_Upper := gIO.i_EL[15].i_ch14,
    sen_Lower := gIO.i_EL[15].i_ch15,
    st_Piston_U_L := stPis_U_L[E_Pis_Name.V4033],
    stOperation := stOper[E_ModeZone.eTank4],
    valve_Upper => gIO.q_EL[4].q_ch15,
    valve_Lower => gIO.q_EL[4].q_ch16); // FB_Piston_U_L
gIO.q_EL[4].q_ch13 := TRUE;

// NETWORK 10
fbPis[E_Pis_Name.V4034](
    sen_Open := gIO.i_EL[16].i_ch3,
    sen_Close := gIO.i_EL[16].i_ch2,
    DefaultCmd := E_PistonDefault_CMD.Close,
    iFB_Num := E_Pis_Name.V4034,
    stOperation := stOper[E_ModeZone.eProduction_Color],
    valve_Open => gIO.q_EL[5].q_ch2); // FB_Piston
fbPis_U_L[E_Pis_Name.V4034](
    enable := fbPis[E_Pis_Name.V4034].valve_Close,
    sen_Upper := gIO.i_EL[16].i_ch4,
    sen_Lower := gIO.i_EL[16].i_ch5,
    st_Piston_U_L := stPis_U_L[E_Pis_Name.V4034],
    stOperation := stOper[E_ModeZone.eTank3],
    valve_Upper => gIO.q_EL[5].q_ch3,
    valve_Lower => gIO.q_EL[5].q_ch4); // FB_Piston_U_L
gIO.q_EL[5].q_ch1 := TRUE;

// NETWORK 11
fbPis[E_Pis_Name.V4035](
    sen_Open := gIO.i_EL[11].i_ch5,
    sen_Close := gIO.i_EL[11].i_ch6,
    DefaultCmd := E_PistonDefault_CMD.Close,
    iFB_Num := E_Pis_Name.V4035,
    stOperation := stOper[E_ModeZone.eProduction_Color],
    valve_Open => gIO.q_Manifold2[16].sol_12); // FB_Piston

// NETWORK 12
fbPis[E_Pis_Name.V4036](
    sen_Open := gIO.i_EL[11].i_ch7,
    sen_Close := gIO.i_EL[11].i_ch8,
    DefaultCmd := E_PistonDefault_CMD.Close,
    iFB_Num := E_Pis_Name.V4036,
    stOperation := stOper[E_ModeZone.eProduction_Color],
    valve_Open => gIO.q_Manifold2[15].sol_12); // FB_Piston

// NETWORK 13
fbPis[E_Pis_Name.V_Dummy_01](
    DefaultCmd := E_PistonDefault_CMD.Close,
    iFB_Num := E_Pis_Name.V_Dummy_01,
    stOperation := stOper[E_ModeZone.eTank1]); // FB_Piston

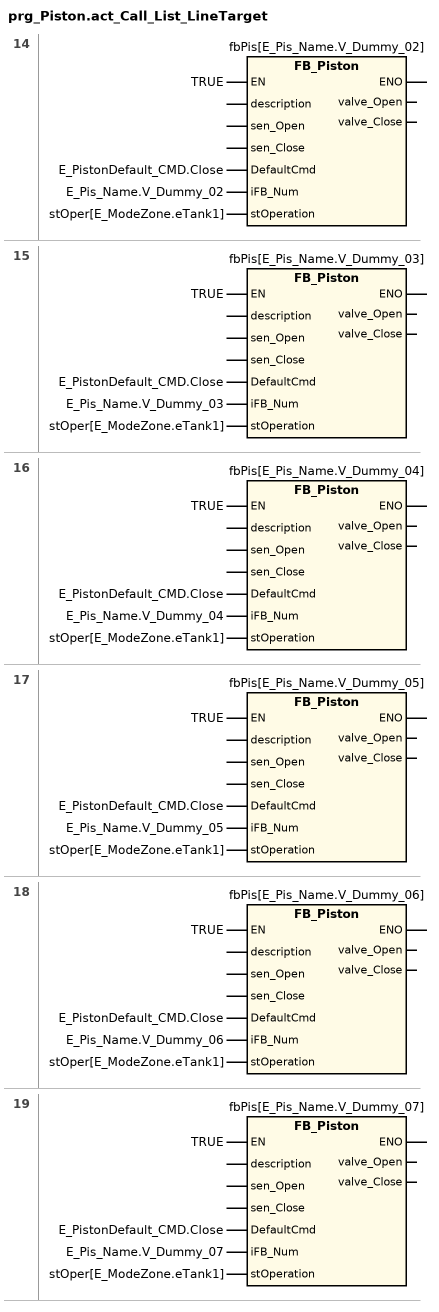
// NETWORK 14
fbPis[E_Pis_Name.V_Dummy_02](
    DefaultCmd := E_PistonDefault_CMD.Close,
    iFB_Num := E_Pis_Name.V_Dummy_02,
    stOperation := stOper[E_ModeZone.eTank1]); // FB_Piston

// NETWORK 15
fbPis[E_Pis_Name.V_Dummy_03](
    DefaultCmd := E_PistonDefault_CMD.Close,
    iFB_Num := E_Pis_Name.V_Dummy_03,
    stOperation := stOper[E_ModeZone.eTank1]); // FB_Piston

// NETWORK 16
fbPis[E_Pis_Name.V_Dummy_04](
    DefaultCmd := E_PistonDefault_CMD.Close,
    iFB_Num := E_Pis_Name.V_Dummy_04,
    stOperation := stOper[E_ModeZone.eTank1]); // FB_Piston

// NETWORK 17
fbPis[E_Pis_Name.V_Dummy_05](
    DefaultCmd := E_PistonDefault_CMD.Close,
    iFB_Num := E_Pis_Name.V_Dummy_05,
    stOperation := stOper[E_ModeZone.eTank1]); // FB_Piston

// NETWORK 18
fbPis[E_Pis_Name.V_Dummy_06](
    DefaultCmd := E_PistonDefault_CMD.Close,
    iFB_Num := E_Pis_Name.V_Dummy_06,
    stOperation := stOper[E_ModeZone.eTank1]); // FB_Piston

// NETWORK 19
fbPis[E_Pis_Name.V_Dummy_07](
    DefaultCmd := E_PistonDefault_CMD.Close,
    iFB_Num := E_Pis_Name.V_Dummy_07,
    stOperation := stOper[E_ModeZone.eTank1]); // FB_Piston

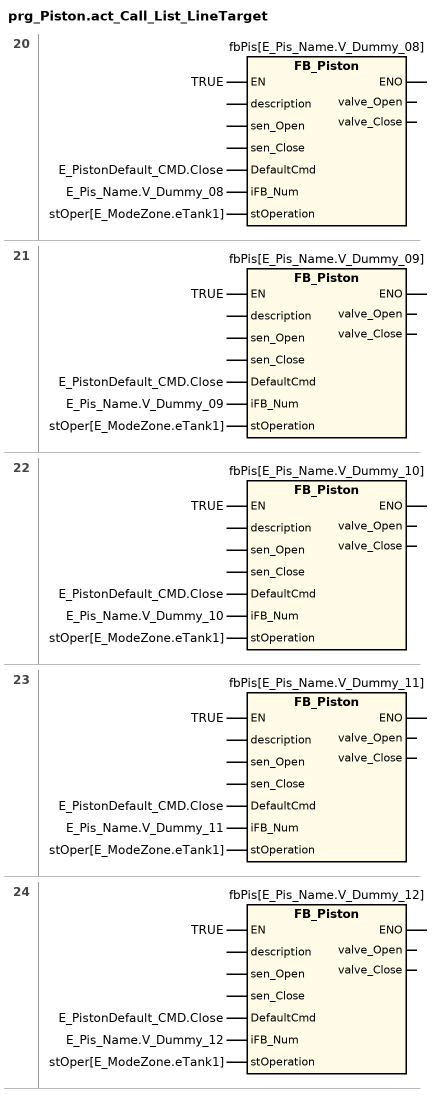
// NETWORK 20
fbPis[E_Pis_Name.V_Dummy_08](
    DefaultCmd := E_PistonDefault_CMD.Close,
    iFB_Num := E_Pis_Name.V_Dummy_08,
    stOperation := stOper[E_ModeZone.eTank1]); // FB_Piston

// NETWORK 21
fbPis[E_Pis_Name.V_Dummy_09](
    DefaultCmd := E_PistonDefault_CMD.Close,
    iFB_Num := E_Pis_Name.V_Dummy_09,
    stOperation := stOper[E_ModeZone.eTank1]); // FB_Piston

// NETWORK 22
fbPis[E_Pis_Name.V_Dummy_10](
    DefaultCmd := E_PistonDefault_CMD.Close,
    iFB_Num := E_Pis_Name.V_Dummy_10,
    stOperation := stOper[E_ModeZone.eTank1]); // FB_Piston

// NETWORK 23
fbPis[E_Pis_Name.V_Dummy_11](
    DefaultCmd := E_PistonDefault_CMD.Close,
    iFB_Num := E_Pis_Name.V_Dummy_11,
    stOperation := stOper[E_ModeZone.eTank1]); // FB_Piston

// NETWORK 24
fbPis[E_Pis_Name.V_Dummy_12](
    DefaultCmd := E_PistonDefault_CMD.Close,
    iFB_Num := E_Pis_Name.V_Dummy_12,
    stOperation := stOper[E_ModeZone.eTank1]); // FB_Piston
END_ACTION

ACTION act_Call_list_TanksColor:
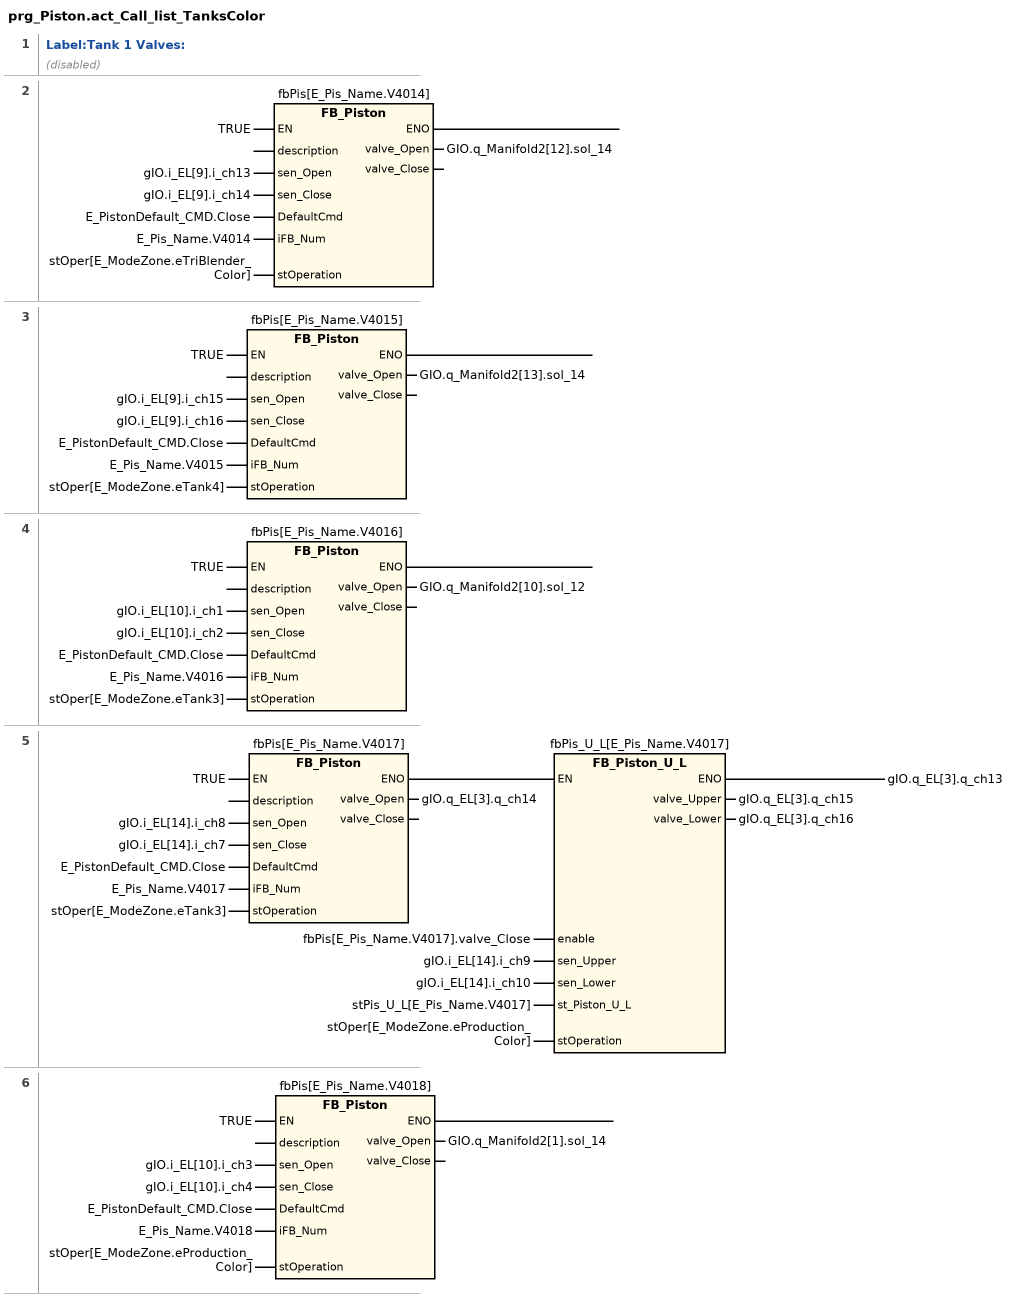
// NETWORK 1 (disabled)
// label: Label:Tank 1 Valves

// NETWORK 2
fbPis[E_Pis_Name.V4014](
    sen_Open := gIO.i_EL[9].i_ch13,
    sen_Close := gIO.i_EL[9].i_ch14,
    DefaultCmd := E_PistonDefault_CMD.Close,
    iFB_Num := E_Pis_Name.V4014,
    stOperation := stOper[E_ModeZone.eTriBlender_Color],
    valve_Open => GIO.q_Manifold2[12].sol_14); // FB_Piston

// NETWORK 3
fbPis[E_Pis_Name.V4015](
    sen_Open := gIO.i_EL[9].i_ch15,
    sen_Close := gIO.i_EL[9].i_ch16,
    DefaultCmd := E_PistonDefault_CMD.Close,
    iFB_Num := E_Pis_Name.V4015,
    stOperation := stOper[E_ModeZone.eTank4],
    valve_Open => GIO.q_Manifold2[13].sol_14); // FB_Piston

// NETWORK 4
fbPis[E_Pis_Name.V4016](
    sen_Open := gIO.i_EL[10].i_ch1,
    sen_Close := gIO.i_EL[10].i_ch2,
    DefaultCmd := E_PistonDefault_CMD.Close,
    iFB_Num := E_Pis_Name.V4016,
    stOperation := stOper[E_ModeZone.eTank3],
    valve_Open => GIO.q_Manifold2[10].sol_12); // FB_Piston

// NETWORK 5
fbPis[E_Pis_Name.V4017](
    sen_Open := gIO.i_EL[14].i_ch8,
    sen_Close := gIO.i_EL[14].i_ch7,
    DefaultCmd := E_PistonDefault_CMD.Close,
    iFB_Num := E_Pis_Name.V4017,
    stOperation := stOper[E_ModeZone.eTank3],
    valve_Open => gIO.q_EL[3].q_ch14); // FB_Piston
fbPis_U_L[E_Pis_Name.V4017](
    enable := fbPis[E_Pis_Name.V4017].valve_Close,
    sen_Upper := gIO.i_EL[14].i_ch9,
    sen_Lower := gIO.i_EL[14].i_ch10,
    st_Piston_U_L := stPis_U_L[E_Pis_Name.V4017],
    stOperation := stOper[E_ModeZone.eProduction_Color],
    valve_Upper => gIO.q_EL[3].q_ch15,
    valve_Lower => gIO.q_EL[3].q_ch16); // FB_Piston_U_L
gIO.q_EL[3].q_ch13 := TRUE;

// NETWORK 6
fbPis[E_Pis_Name.V4018](
    sen_Open := gIO.i_EL[10].i_ch3,
    sen_Close := gIO.i_EL[10].i_ch4,
    DefaultCmd := E_PistonDefault_CMD.Close,
    iFB_Num := E_Pis_Name.V4018,
    stOperation := stOper[E_ModeZone.eProduction_Color],
    valve_Open => GIO.q_Manifold2[1].sol_14); // FB_Piston

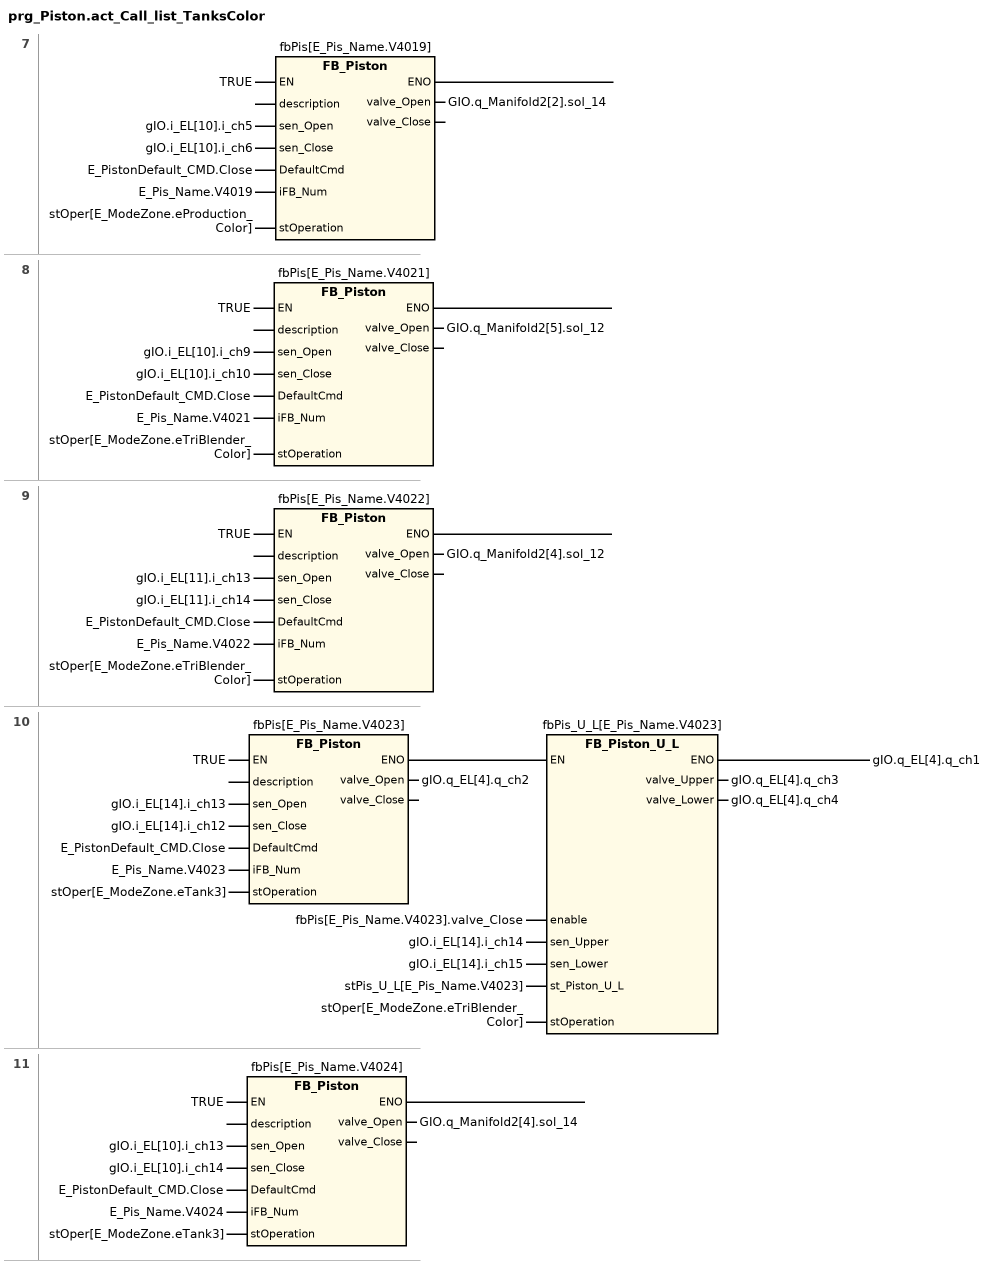
// NETWORK 7
fbPis[E_Pis_Name.V4019](
    sen_Open := gIO.i_EL[10].i_ch5,
    sen_Close := gIO.i_EL[10].i_ch6,
    DefaultCmd := E_PistonDefault_CMD.Close,
    iFB_Num := E_Pis_Name.V4019,
    stOperation := stOper[E_ModeZone.eProduction_Color],
    valve_Open => GIO.q_Manifold2[2].sol_14); // FB_Piston

// NETWORK 8
fbPis[E_Pis_Name.V4021](
    sen_Open := gIO.i_EL[10].i_ch9,
    sen_Close := gIO.i_EL[10].i_ch10,
    DefaultCmd := E_PistonDefault_CMD.Close,
    iFB_Num := E_Pis_Name.V4021,
    stOperation := stOper[E_ModeZone.eTriBlender_Color],
    valve_Open => GIO.q_Manifold2[5].sol_12); // FB_Piston

// NETWORK 9
fbPis[E_Pis_Name.V4022](
    sen_Open := gIO.i_EL[11].i_ch13,
    sen_Close := gIO.i_EL[11].i_ch14,
    DefaultCmd := E_PistonDefault_CMD.Close,
    iFB_Num := E_Pis_Name.V4022,
    stOperation := stOper[E_ModeZone.eTriBlender_Color],
    valve_Open => GIO.q_Manifold2[4].sol_12); // FB_Piston

// NETWORK 10
fbPis[E_Pis_Name.V4023](
    sen_Open := gIO.i_EL[14].i_ch13,
    sen_Close := gIO.i_EL[14].i_ch12,
    DefaultCmd := E_PistonDefault_CMD.Close,
    iFB_Num := E_Pis_Name.V4023,
    stOperation := stOper[E_ModeZone.eTank3],
    valve_Open => gIO.q_EL[4].q_ch2); // FB_Piston
fbPis_U_L[E_Pis_Name.V4023](
    enable := fbPis[E_Pis_Name.V4023].valve_Close,
    sen_Upper := gIO.i_EL[14].i_ch14,
    sen_Lower := gIO.i_EL[14].i_ch15,
    st_Piston_U_L := stPis_U_L[E_Pis_Name.V4023],
    stOperation := stOper[E_ModeZone.eTriBlender_Color],
    valve_Upper => gIO.q_EL[4].q_ch3,
    valve_Lower => gIO.q_EL[4].q_ch4); // FB_Piston_U_L
gIO.q_EL[4].q_ch1 := TRUE;

// NETWORK 11
fbPis[E_Pis_Name.V4024](
    sen_Open := gIO.i_EL[10].i_ch13,
    sen_Close := gIO.i_EL[10].i_ch14,
    DefaultCmd := E_PistonDefault_CMD.Close,
    iFB_Num := E_Pis_Name.V4024,
    stOperation := stOper[E_ModeZone.eTank3],
    valve_Open => GIO.q_Manifold2[4].sol_14); // FB_Piston

